// I:1800 (MONETcommon#17): a slew still running after 600 s is software error 16#40 and the slew is dropped. The time seam divides every
// timeout by 1000, so the 600 s are 0.6 s; the mock move takes far longer.
METHOD PRIVATE Slew_Times_Out_After_600_Seconds
VAR_INST
	rig			: FB_IagRig;
	nStep		: INT;
	nCycles		: UINT;
	sTest		: STRING(80);
END_VAR
TEST('Slew_Times_Out_After_600_Seconds');
sTest := 'Slew_Times_Out_After_600_Seconds: ';
IF nStep >= 90 THEN
	RETURN;
END_IF
rig.Scan();
nCycles := nCycles + 1;
CASE nStep OF
0:	// wait for the clock, then power on
	IF rig.ClockValid THEN
		rig.fbTel.Init();
		nStep := 10;
		nCycles := 0;
	ELSIF nCycles > 2000 THEN
		AssertTrue(Condition := FALSE, Message := 'the astronomical clock never became valid');
		F_Note(bFailed := TRUE, sText := CONCAT(sTest, 'the astronomical clock never became valid'));
		rig.SetTimeDivisor(nValue := 1);
		nStep := 99;
		TEST_FINISHED();
	END_IF
10:	IF rig.Online THEN
		rig.SetMoveScans(nScans := 60000);
		rig.SetTimeDivisor(nValue := 1000);
		rig.fbTel.Slew(fAzimuth := 180.0, fAltitude := 45.0);
		nStep := 20;
		nCycles := 0;
	ELSIF nCycles > 1500 THEN
		AssertTrue(Condition := FALSE, Message := 'the mock telescope did not reach READY_STATE 1.0');
		F_Note(bFailed := TRUE, sText := CONCAT(sTest, 'the mock telescope did not reach READY_STATE 1.0'));
		rig.SetTimeDivisor(nValue := 1);
		nStep := 99;
		TEST_FINISHED();
	END_IF
20:
	IF rig.fbTel.bError THEN
		AssertTrue(Condition := rig.fbTel.bSoftwareError AND rig.fbTel.nSoftwareErrorID = 16#40, Message := 'the slew timeout is software error 16#40');
		F_Note(bFailed := NOT (rig.fbTel.bSoftwareError AND rig.fbTel.nSoftwareErrorID = 16#40), sText := CONCAT(sTest, 'the slew timeout is software error 16#40'));
		AssertTrue(Condition := NOT rig.fbTel.bSlewActive, Message := 'the slew is dropped');
		F_Note(bFailed := NOT (NOT rig.fbTel.bSlewActive), sText := CONCAT(sTest, 'the slew is dropped'));
		rig.SetTimeDivisor(nValue := 1);
		nStep := 99;
		TEST_FINISHED();
	ELSIF nCycles > 3000 THEN
		AssertTrue(Condition := FALSE, Message := 'the slew never timed out');
		F_Note(bFailed := TRUE, sText := CONCAT(sTest, 'the slew never timed out'));
		rig.SetTimeDivisor(nValue := 1);
		nStep := 99;
		TEST_FINISHED();
	END_IF
END_CASE
END_METHOD

// I:466, 491-496: an online telescope without a command for 12 h parks itself (tonPowerTimeout). The time seam divides by 1000000, so the
// 12 h are 43 ms.
METHOD PRIVATE Idle_Telescope_Parks_After_12_Hours
VAR_INST
	rig			: FB_IagRig;
	nStep		: INT;
	nCycles		: UINT;
	sTest		: STRING(80);
END_VAR
TEST('Idle_Telescope_Parks_After_12_Hours');
sTest := 'Idle_Telescope_Parks_After_12_Hours: ';
IF nStep >= 90 THEN
	RETURN;
END_IF
rig.Scan();
nCycles := nCycles + 1;
CASE nStep OF
0:	// wait for the clock, then power on
	IF rig.ClockValid THEN
		rig.fbTel.Init();
		nStep := 10;
		nCycles := 0;
	ELSIF nCycles > 2000 THEN
		AssertTrue(Condition := FALSE, Message := 'the astronomical clock never became valid');
		F_Note(bFailed := TRUE, sText := CONCAT(sTest, 'the astronomical clock never became valid'));
		rig.SetTimeDivisor(nValue := 1);
		nStep := 99;
		TEST_FINISHED();
	END_IF
10:	IF rig.Online THEN
		rig.SetTimeDivisor(nValue := 1000000);
		nStep := 20;
		nCycles := 0;
	ELSIF nCycles > 1500 THEN
		AssertTrue(Condition := FALSE, Message := 'the mock telescope did not reach READY_STATE 1.0');
		F_Note(bFailed := TRUE, sText := CONCAT(sTest, 'the mock telescope did not reach READY_STATE 1.0'));
		rig.SetTimeDivisor(nValue := 1);
		nStep := 99;
		TEST_FINISHED();
	END_IF
20:
	IF rig.fbTel.bParkActive OR rig.fbTel.bIsParked THEN
		rig.SetTimeDivisor(nValue := 1);
		AssertTrue(Condition := rig.fbTel.bParkActive OR rig.fbTel.bIsParked, Message := 'the idle telescope parked itself');
		F_Note(bFailed := NOT (rig.fbTel.bParkActive OR rig.fbTel.bIsParked), sText := CONCAT(sTest, 'the idle telescope parked itself'));
		nStep := 99;
		TEST_FINISHED();
	ELSIF nCycles > 3000 THEN
		AssertTrue(Condition := FALSE, Message := 'the idle telescope never parked');
		F_Note(bFailed := TRUE, sText := CONCAT(sTest, 'the idle telescope never parked'));
		rig.SetTimeDivisor(nValue := 1);
		nStep := 99;
		TEST_FINISHED();
	END_IF
END_CASE
END_METHOD

END_FUNCTION_BLOCK

// ---- POUs/IagParkDuringPowerOn_Tests.TcPOU
// Characterization of FB_TelescopeControl (IAG50cm) for a park or a stop that arrives during the power-on, on mock axes (plan step 2,
// IAG50cmTests README). These tests pin what the code does today, with the line of the behaviour in a comment; they are not a
// specification. Every test owns a rig and runs over many PLC cycles (VAR_INST of the method, one Scan() per cycle). Failed checks
// are also noted in GVL_Diag.sFailures (printed by Run-Tests.ps1).
FUNCTION_BLOCK IagParkDuringPowerOn_Tests EXTENDS TcUnit.FB_TestSuite
VAR
END_VAR

Park_During_PowerOn_Aborts_The_Startup_And_Parks();
Stop_During_PowerOn_Aborts_The_Startup();
AxesOff_Park_After_Stopped_Startup_Reports_Parked();
AxesOff_Park_With_Slow_Covers_Reports_Parking_Then_Parked();
Stop_During_AxesOff_Park_Does_Not_Cancel_It();
AxesOff_Park_Gives_Up_When_The_Covers_Do_Not_Close();
Park_In_The_Sweep_Parks_In_Place();
Park_After_Stage_100_Still_Moves_To_The_Park_Position();

// I:529-541 (IAG50cm#109): a park that arrives while the power-on runs outranks it, like a stop: the startup is aborted, the
// covers the power-on opened are closed again and the telescope ends parked, never ready (READY_STATE does not reach 1.0).
// In the covers phase the axes are still off, so the park takes the axes-off path (#54, #110): covers closed, dome parked,
// the mount is not moved, READY_STATE 0.0 and bIsParked is TRUE with bParkedInPlace (#187). Decision 3 of the plan: as MONET (MONETcommon#87).
METHOD PRIVATE Park_During_PowerOn_Aborts_The_Startup_And_Parks
VAR_INST
	rig			: FB_IagRig;
	nStep		: INT;
	nCycles		: UINT;
	sTest		: STRING(80);
END_VAR
TEST('Park_During_PowerOn_Aborts_The_Startup_And_Parks');
sTest := 'Park_During_PowerOn_Aborts_The_Startup_And_Parks: ';
IF nStep >= 90 THEN
	RETURN;
END_IF
rig.Scan();
nCycles := nCycles + 1;
CASE nStep OF
0:	// wait for the clock, then power on
	IF rig.ClockValid THEN
		rig.fbTel.Init();
		nStep := 10;
		nCycles := 0;
	ELSIF nCycles > 2000 THEN
		AssertTrue(Condition := FALSE, Message := 'the astronomical clock never became valid');
		F_Note(bFailed := TRUE, sText := CONCAT(sTest, 'the astronomical clock never became valid'));
		nStep := 99;
		TEST_FINISHED();
	END_IF
10:	// the power-on has commanded the covers: park now
	IF rig.fbCovers.nOpenCalls >= 1 THEN
		rig.fbTel.Park();
		nStep := 20;
		nCycles := 0;
	ELSIF nCycles > 300 THEN
		AssertTrue(Condition := FALSE, Message := 'the power-on never commanded the covers');
		F_Note(bFailed := TRUE, sText := CONCAT(sTest, 'the power-on never commanded the covers'));
		nStep := 99;
		TEST_FINISHED();
	END_IF
20:	// the power-on is aborted at once, the covers are commanded closed
	IF nCycles = 3 THEN
		AssertTrue(Condition := NOT rig.fbTel.bPowerActive, Message := 'the power-on is aborted');
		F_Note(bFailed := (rig.fbTel.bPowerActive), sText := CONCAT(sTest, 'the power-on is aborted'));
		nStep := 30;
		nCycles := 0;
	END_IF
30:	// the park finishes (READY_STATE 0.0, the axes were off: bIsParked TRUE with bParkedInPlace, #187), the startup never does
	AssertFalse(Condition := rig.Online, Message := 'the startup went on to the end');
	F_Note(bFailed := (rig.Online), sText := CONCAT(sTest, 'the startup went on to the end'));
	IF rig.fbTel.ReadyState = 0.0 THEN
		AssertTrue(Condition := rig.fbCovers.nCloseCalls >= 1, Message := 'the covers were closed');
		F_Note(bFailed := NOT (rig.fbCovers.nCloseCalls >= 1), sText := CONCAT(sTest, 'the covers were closed'));
		AssertTrue(Condition := rig.fbTel.bIsParked, Message := 'bIsParked is TRUE (#187)');
		F_Note(bFailed := NOT (rig.fbTel.bIsParked), sText := CONCAT(sTest, 'bIsParked is TRUE (#187)'));
		AssertTrue(Condition := rig.fbTel.bParkedInPlace, Message := 'bParkedInPlace is TRUE, the mount was not moved');
		F_Note(bFailed := NOT (rig.fbTel.bParkedInPlace), sText := CONCAT(sTest, 'bParkedInPlace is TRUE, the mount was not moved'));
		nStep := 99;
		TEST_FINISHED();
	ELSIF nCycles > 1500 THEN
		AssertTrue(Condition := FALSE, Message := 'the telescope did not park');
		F_Note(bFailed := TRUE, sText := CONCAT(sTest, 'the telescope did not park'));
		nStep := 99;
		TEST_FINISHED();
	END_IF
END_CASE
END_METHOD

// I:501-526 (#27): an explicit stop outranks the power-on: the startup is aborted (READY_STATE -2.0), nothing is parked and the
// covers the power-on opened stay open.
METHOD PRIVATE Stop_During_PowerOn_Aborts_The_Startup
VAR_INST
	rig			: FB_IagRig;
	nStep		: INT;
	nCycles		: UINT;
	sTest		: STRING(80);
END_VAR
TEST('Stop_During_PowerOn_Aborts_The_Startup');
sTest := 'Stop_During_PowerOn_Aborts_The_Startup: ';
IF nStep >= 90 THEN
	RETURN;
END_IF
rig.Scan();
nCycles := nCycles + 1;
CASE nStep OF
0:	// wait for the clock, then power on
	IF rig.ClockValid THEN
		rig.fbTel.Init();
		nStep := 10;
		nCycles := 0;
	ELSIF nCycles > 2000 THEN
		AssertTrue(Condition := FALSE, Message := 'the astronomical clock never became valid');
		F_Note(bFailed := TRUE, sText := CONCAT(sTest, 'the astronomical clock never became valid'));
		nStep := 99;
		TEST_FINISHED();
	END_IF
10:	// the power-on has commanded the covers: stop now
	IF rig.fbCovers.nOpenCalls >= 1 THEN
		rig.fbTel.Stop();
		nStep := 20;
		nCycles := 0;
	ELSIF nCycles > 300 THEN
		AssertTrue(Condition := FALSE, Message := 'the power-on never commanded the covers');
		F_Note(bFailed := TRUE, sText := CONCAT(sTest, 'the power-on never commanded the covers'));
		nStep := 99;
		TEST_FINISHED();
	END_IF
20:	// wait until the stop has settled
	IF NOT rig.fbTel.bStopActive AND rig.fbTel.bStopped AND nCycles > 5 THEN
		AssertFalse(Condition := rig.fbTel.bPowerActive, Message := 'the power-on request is dropped');
		F_Note(bFailed := (rig.fbTel.bPowerActive), sText := CONCAT(sTest, 'the power-on request is dropped'));
		AssertFalse(Condition := rig.fbTel.bParkActive OR rig.fbTel.bIsParked, Message := 'the stop does not park');
		F_Note(bFailed := (rig.fbTel.bParkActive OR rig.fbTel.bIsParked), sText := CONCAT(sTest, 'the stop does not park'));
		AssertTrue(Condition := rig.fbTel.ReadyState = -2.0, Message := 'READY_STATE is -2.0 (startup aborted)');
		F_Note(bFailed := NOT (rig.fbTel.ReadyState = -2.0), sText := CONCAT(sTest, 'READY_STATE is -2.0 (startup aborted)'));
		AssertTrue(Condition := rig.fbCovers.nCloseCalls = 0 AND rig.fbCovers.bOpened, Message := 'the covers stay open');
		F_Note(bFailed := NOT (rig.fbCovers.nCloseCalls = 0 AND rig.fbCovers.bOpened), sText := CONCAT(sTest, 'the covers stay open'));
		nStep := 99;
		TEST_FINISHED();
	ELSIF nCycles > 400 THEN
		AssertTrue(Condition := FALSE, Message := 'the stop did not settle');
		F_Note(bFailed := TRUE, sText := CONCAT(sTest, 'the stop did not settle'));
		nStep := 99;
		TEST_FINISHED();
	END_IF
END_CASE
END_METHOD

// IAG50cm#110: after a stopped startup (-2) a park with the axes off closes the covers and parks the dome, the mount is not moved.
// READY_STATE leaves -2 for 0.0 and bIsParked becomes TRUE with bParkedInPlace (#187); a new power-on clears both.
METHOD PRIVATE AxesOff_Park_After_Stopped_Startup_Reports_Parked
VAR_INST
	rig			: FB_IagRig;
	nStep		: INT;
	nCycles		: UINT;
	sTest		: STRING(80);
END_VAR
TEST('AxesOff_Park_After_Stopped_Startup_Reports_Parked');
sTest := 'AxesOff_Park_After_Stopped_Startup_Reports_Parked: ';
IF nStep >= 90 THEN
	RETURN;
END_IF
rig.Scan();
nCycles := nCycles + 1;
CASE nStep OF
0:	// wait for the clock, then power on
	IF rig.ClockValid THEN
		rig.fbTel.Init();
		nStep := 10;
		nCycles := 0;
	ELSIF nCycles > 2000 THEN
		AssertTrue(Condition := FALSE, Message := 'the astronomical clock never became valid');
		F_Note(bFailed := TRUE, sText := CONCAT(sTest, 'the astronomical clock never became valid'));
		nStep := 99;
		TEST_FINISHED();
	END_IF
10:	// the power-on has commanded the covers: stop now
	IF rig.fbCovers.nOpenCalls >= 1 THEN
		rig.fbTel.Stop();
		nStep := 20;
		nCycles := 0;
	ELSIF nCycles > 300 THEN
		AssertTrue(Condition := FALSE, Message := 'the power-on never commanded the covers');
		F_Note(bFailed := TRUE, sText := CONCAT(sTest, 'the power-on never commanded the covers'));
		nStep := 99;
		TEST_FINISHED();
	END_IF
20:	// the stop has settled: -2, then park with the axes off
	IF NOT rig.fbTel.bStopActive AND rig.fbTel.bStopped AND nCycles > 5 THEN
		AssertTrue(Condition := rig.fbTel.ReadyState = -2.0, Message := 'READY_STATE is -2.0 after the stop');
		F_Note(bFailed := NOT (rig.fbTel.ReadyState = -2.0), sText := CONCAT(sTest, 'READY_STATE is -2.0 after the stop'));
		rig.fbTel.Park();
		nStep := 30;
		nCycles := 0;
	ELSIF nCycles > 400 THEN
		AssertTrue(Condition := FALSE, Message := 'the stop did not settle');
		F_Note(bFailed := TRUE, sText := CONCAT(sTest, 'the stop did not settle'));
		nStep := 99;
		TEST_FINISHED();
	END_IF
30:	// the covers close, READY_STATE becomes 0.0, bIsParked is TRUE (#187)
	IF rig.fbTel.ReadyState = 0.0 THEN
		AssertTrue(Condition := rig.fbCovers.nCloseCalls >= 1, Message := 'the covers were closed');
		F_Note(bFailed := NOT (rig.fbCovers.nCloseCalls >= 1), sText := CONCAT(sTest, 'the covers were closed'));
		AssertTrue(Condition := rig.fbTel.bIsParked, Message := 'bIsParked is TRUE (#187)');
		F_Note(bFailed := NOT (rig.fbTel.bIsParked), sText := CONCAT(sTest, 'bIsParked is TRUE (#187)'));
		AssertTrue(Condition := rig.fbTel.bParkedInPlace, Message := 'bParkedInPlace is TRUE, the mount was not moved');
		F_Note(bFailed := NOT (rig.fbTel.bParkedInPlace), sText := CONCAT(sTest, 'bParkedInPlace is TRUE, the mount was not moved'));
		rig.fbTel.Init();
		nStep := 40;
		nCycles := 0;
	ELSIF nCycles > 400 THEN
		AssertTrue(Condition := FALSE, Message := 'READY_STATE did not reach 0.0');
		F_Note(bFailed := TRUE, sText := CONCAT(sTest, 'READY_STATE did not reach 0.0'));
		nStep := 99;
		TEST_FINISHED();
	END_IF
40:	// a new power-on ends the covered state
	IF rig.fbTel.ReadyState > 0.0 THEN
		nStep := 99;
		TEST_FINISHED();
	ELSIF nCycles > 400 THEN
		AssertTrue(Condition := FALSE, Message := 'the new power-on did not leave READY_STATE 0.0');
		F_Note(bFailed := TRUE, sText := CONCAT(sTest, 'the new power-on did not leave READY_STATE 0.0'));
		nStep := 99;
		TEST_FINISHED();
	END_IF
END_CASE
END_METHOD

// IAG50cm#187: an axes-off park whose covers close slowly reports READY_STATE 0.3 and bIsParked FALSE while they are open, and
// parked in place (READY_STATE 0.0, bIsParked and bParkedInPlace TRUE) once they are closed. The covers mock holds the close.
METHOD PRIVATE AxesOff_Park_With_Slow_Covers_Reports_Parking_Then_Parked
VAR_INST
	rig			: FB_IagRig;
	nStep		: INT;
	nCycles		: UINT;
	sTest		: STRING(80);
END_VAR
TEST('AxesOff_Park_With_Slow_Covers_Reports_Parking_Then_Parked');
sTest := 'AxesOff_Park_With_Slow_Covers_Reports_Parking_Then_Parked: ';
IF nStep >= 90 THEN
	RETURN;
END_IF
rig.Scan();
nCycles := nCycles + 1;
CASE nStep OF
0:	// wait for the clock, then power on
	IF rig.ClockValid THEN
		rig.fbTel.Init();
		nStep := 10;
		nCycles := 0;
	ELSIF nCycles > 2000 THEN
		AssertTrue(Condition := FALSE, Message := 'the astronomical clock never became valid');
		F_Note(bFailed := TRUE, sText := CONCAT(sTest, 'the astronomical clock never became valid'));
		nStep := 99;
		TEST_FINISHED();
	END_IF
10:	// the power-on has commanded the covers: stop now
	IF rig.fbCovers.nOpenCalls >= 1 THEN
		rig.fbTel.Stop();
		nStep := 20;
		nCycles := 0;
	ELSIF nCycles > 300 THEN
		AssertTrue(Condition := FALSE, Message := 'the power-on never commanded the covers');
		F_Note(bFailed := TRUE, sText := CONCAT(sTest, 'the power-on never commanded the covers'));
		nStep := 99;
		TEST_FINISHED();
	END_IF
20:	// the stop has settled: the covers now close slowly, park with the axes off
	IF NOT rig.fbTel.bStopActive AND rig.fbTel.bStopped AND nCycles > 5 THEN
		rig.fbCovers.HoldClose(bHold := TRUE);
		rig.fbTel.Park();
		nStep := 30;
		nCycles := 0;
	ELSIF nCycles > 400 THEN
		AssertTrue(Condition := FALSE, Message := 'the stop did not settle');
		F_Note(bFailed := TRUE, sText := CONCAT(sTest, 'the stop did not settle'));
		nStep := 99;
		TEST_FINISHED();
	END_IF
30:	// the covers were commanded but are not closed: 0.3 (parking), not parked, not 0 and not -2
	IF rig.fbCovers.nCloseCalls >= 1 AND nCycles > 20 THEN
		AssertTrue(Condition := rig.fbTel.ReadyState = 0.3, Message := 'READY_STATE is 0.3 while the covers close (#187)');
		F_Note(bFailed := NOT (rig.fbTel.ReadyState = 0.3), sText := CONCAT(sTest, 'READY_STATE is 0.3 while the covers close (#187)'));
		AssertTrue(Condition := NOT rig.fbTel.bIsParked, Message := 'bIsParked stays FALSE until the covers are closed');
		F_Note(bFailed := NOT (NOT rig.fbTel.bIsParked), sText := CONCAT(sTest, 'bIsParked stays FALSE until the covers are closed'));
		AssertTrue(Condition := rig.fbTel.bSafeParked, Message := 'the axes-off park is pending');
		F_Note(bFailed := NOT (rig.fbTel.bSafeParked), sText := CONCAT(sTest, 'the axes-off park is pending'));
		rig.fbCovers.FinishClose();
		nStep := 40;
		nCycles := 0;
	ELSIF nCycles > 400 THEN
		AssertTrue(Condition := FALSE, Message := 'the covers were never commanded to close');
		F_Note(bFailed := TRUE, sText := CONCAT(sTest, 'the covers were never commanded to close'));
		nStep := 99;
		TEST_FINISHED();
	END_IF
40:	// the covers closed: parked in place
	IF rig.fbTel.ReadyState = 0.0 THEN
		AssertTrue(Condition := rig.fbTel.bIsParked, Message := 'bIsParked is TRUE once the covers are closed (#187)');
		F_Note(bFailed := NOT (rig.fbTel.bIsParked), sText := CONCAT(sTest, 'bIsParked is TRUE once the covers are closed (#187)'));
		AssertTrue(Condition := rig.fbTel.bParkedInPlace, Message := 'bParkedInPlace is TRUE, the mount was not moved');
		F_Note(bFailed := NOT (rig.fbTel.bParkedInPlace), sText := CONCAT(sTest, 'bParkedInPlace is TRUE, the mount was not moved'));
		AssertTrue(Condition := NOT rig.fbTel.bSafeParked, Message := 'the axes-off park is finished');
		F_Note(bFailed := NOT (NOT rig.fbTel.bSafeParked), sText := CONCAT(sTest, 'the axes-off park is finished'));
		nStep := 99;
		TEST_FINISHED();
	ELSIF nCycles > 400 THEN
		AssertTrue(Condition := FALSE, Message := 'READY_STATE did not reach 0.0 after the covers closed');
		F_Note(bFailed := TRUE, sText := CONCAT(sTest, 'READY_STATE did not reach 0.0 after the covers closed'));
		nStep := 99;
		TEST_FINISHED();
	END_IF
END_CASE
END_METHOD

// IAG50cm#196: a stop during the axes-off park (covers closing) is ignored and logged ('Stop ignored'): the park goes on and ends parked in place.
METHOD PRIVATE Stop_During_AxesOff_Park_Does_Not_Cancel_It
VAR_INST
	rig			: FB_IagRig;
	nStep		: INT;
	nCycles		: UINT;
	sTest		: STRING(80);
END_VAR
TEST('Stop_During_AxesOff_Park_Does_Not_Cancel_It');
sTest := 'Stop_During_AxesOff_Park_Does_Not_Cancel_It: ';
IF nStep >= 90 THEN
	RETURN;
END_IF
rig.Scan();
nCycles := nCycles + 1;
CASE nStep OF
0:	// wait for the clock, then power on
	IF rig.ClockValid THEN
		rig.fbTel.Init();
		nStep := 10;
		nCycles := 0;
	ELSIF nCycles > 2000 THEN
		AssertTrue(Condition := FALSE, Message := 'the astronomical clock never became valid');
		F_Note(bFailed := TRUE, sText := CONCAT(sTest, 'the astronomical clock never became valid'));
		nStep := 99;
		TEST_FINISHED();
	END_IF
10:	// the power-on has commanded the covers: stop now
	IF rig.fbCovers.nOpenCalls >= 1 THEN
		rig.fbTel.Stop();
		nStep := 20;
		nCycles := 0;
	ELSIF nCycles > 300 THEN
		AssertTrue(Condition := FALSE, Message := 'the power-on never commanded the covers');
		F_Note(bFailed := TRUE, sText := CONCAT(sTest, 'the power-on never commanded the covers'));
		nStep := 99;
		TEST_FINISHED();
	END_IF
20:	// the stop has settled: the covers now close slowly, park with the axes off
	IF NOT rig.fbTel.bStopActive AND rig.fbTel.bStopped AND nCycles > 5 THEN
		rig.fbCovers.HoldClose(bHold := TRUE);
		rig.fbTel.Park();
		nStep := 30;
		nCycles := 0;
	ELSIF nCycles > 400 THEN
		AssertTrue(Condition := FALSE, Message := 'the stop did not settle');
		F_Note(bFailed := TRUE, sText := CONCAT(sTest, 'the stop did not settle'));
		nStep := 99;
		TEST_FINISHED();
	END_IF
30:	// the covers were commanded but are not closed: 0.3 (parking), not parked, not 0 and not -2
	IF rig.fbCovers.nCloseCalls >= 1 AND nCycles > 20 THEN
		AssertTrue(Condition := rig.fbTel.ReadyState = 0.3, Message := 'READY_STATE is 0.3 while the covers close (#187)');
		F_Note(bFailed := NOT (rig.fbTel.ReadyState = 0.3), sText := CONCAT(sTest, 'READY_STATE is 0.3 while the covers close (#187)'));
		AssertTrue(Condition := NOT rig.fbTel.bIsParked, Message := 'bIsParked stays FALSE until the covers are closed');
		F_Note(bFailed := NOT (NOT rig.fbTel.bIsParked), sText := CONCAT(sTest, 'bIsParked stays FALSE until the covers are closed'));
		AssertTrue(Condition := rig.fbTel.bSafeParked, Message := 'the axes-off park is pending');
		F_Note(bFailed := NOT (rig.fbTel.bSafeParked), sText := CONCAT(sTest, 'the axes-off park is pending'));
		rig.fbTel.Stop();
		nStep := 35;
		nCycles := 0;
	ELSIF nCycles > 400 THEN
		AssertTrue(Condition := FALSE, Message := 'the covers were never commanded to close');
		F_Note(bFailed := TRUE, sText := CONCAT(sTest, 'the covers were never commanded to close'));
		nStep := 99;
		TEST_FINISHED();
	END_IF
35:	// the stop has settled: the park was not cancelled
	IF NOT rig.fbTel.bStopActive AND nCycles > 5 THEN
		AssertTrue(Condition := rig.fbTel.bSafeParked, Message := 'the stop does not cancel the axes-off park (#196)');
		F_Note(bFailed := NOT (rig.fbTel.bSafeParked), sText := CONCAT(sTest, 'the stop does not cancel the axes-off park (#196)'));
		AssertTrue(Condition := rig.fbTel.ReadyState = 0.3, Message := 'READY_STATE stays 0.3 after the stop (#196)');
		F_Note(bFailed := NOT (rig.fbTel.ReadyState = 0.3), sText := CONCAT(sTest, 'READY_STATE stays 0.3 after the stop (#196)'));
		rig.fbCovers.FinishClose();
		nStep := 40;
		nCycles := 0;
	ELSIF nCycles > 400 THEN
		AssertTrue(Condition := FALSE, Message := 'the stop did not settle');
		F_Note(bFailed := TRUE, sText := CONCAT(sTest, 'the stop did not settle'));
		nStep := 99;
		TEST_FINISHED();
	END_IF
40:	// the covers closed: parked in place
	IF rig.fbTel.ReadyState = 0.0 THEN
		AssertTrue(Condition := rig.fbTel.bIsParked, Message := 'bIsParked is TRUE once the covers are closed (#187)');
		F_Note(bFailed := NOT (rig.fbTel.bIsParked), sText := CONCAT(sTest, 'bIsParked is TRUE once the covers are closed (#187)'));
		AssertTrue(Condition := rig.fbTel.bParkedInPlace, Message := 'bParkedInPlace is TRUE, the mount was not moved');
		F_Note(bFailed := NOT (rig.fbTel.bParkedInPlace), sText := CONCAT(sTest, 'bParkedInPlace is TRUE, the mount was not moved'));
		AssertTrue(Condition := NOT rig.fbTel.bSafeParked, Message := 'the axes-off park is finished');
		F_Note(bFailed := NOT (NOT rig.fbTel.bSafeParked), sText := CONCAT(sTest, 'the axes-off park is finished'));
		nStep := 99;
		TEST_FINISHED();
	ELSIF nCycles > 400 THEN
		AssertTrue(Condition := FALSE, Message := 'READY_STATE did not reach 0.0 after the covers closed');
		F_Note(bFailed := TRUE, sText := CONCAT(sTest, 'READY_STATE did not reach 0.0 after the covers closed'));
		nStep := 99;
		TEST_FINISHED();
	END_IF
END_CASE
END_METHOD

// IAG50cm#187: an axes-off park whose covers never close gives up after 120 s (the time seam divides by 1000): bSafeParked is dropped,
// READY_STATE is not 0.3 for ever and the telescope is never reported parked.
METHOD PRIVATE AxesOff_Park_Gives_Up_When_The_Covers_Do_Not_Close
VAR_INST
	rig			: FB_IagRig;
	nStep		: INT;
	nCycles		: UINT;
	sTest		: STRING(80);
END_VAR
TEST('AxesOff_Park_Gives_Up_When_The_Covers_Do_Not_Close');
sTest := 'AxesOff_Park_Gives_Up_When_The_Covers_Do_Not_Close: ';
IF nStep >= 90 THEN
	RETURN;
END_IF
rig.Scan();
nCycles := nCycles + 1;
CASE nStep OF
0:	// wait for the clock, then power on
	IF rig.ClockValid THEN
		rig.fbTel.Init();
		nStep := 10;
		nCycles := 0;
	ELSIF nCycles > 2000 THEN
		AssertTrue(Condition := FALSE, Message := 'the astronomical clock never became valid');
		F_Note(bFailed := TRUE, sText := CONCAT(sTest, 'the astronomical clock never became valid'));
		nStep := 99;
		TEST_FINISHED();
	END_IF
10:	// the power-on has commanded the covers: stop now
	IF rig.fbCovers.nOpenCalls >= 1 THEN
		rig.fbTel.Stop();
		nStep := 20;
		nCycles := 0;
	ELSIF nCycles > 300 THEN
		AssertTrue(Condition := FALSE, Message := 'the power-on never commanded the covers');
		F_Note(bFailed := TRUE, sText := CONCAT(sTest, 'the power-on never commanded the covers'));
		nStep := 99;
		TEST_FINISHED();
	END_IF
20:	// the stop has settled: the covers never close, park with the axes off; 120 s are 0.12 s
	IF NOT rig.fbTel.bStopActive AND rig.fbTel.bStopped AND nCycles > 5 THEN
		rig.fbCovers.HoldClose(bHold := TRUE);
		rig.SetTimeDivisor(nValue := 1000);
		rig.fbTel.Park();
		nStep := 30;
		nCycles := 0;
	ELSIF nCycles > 400 THEN
		AssertTrue(Condition := FALSE, Message := 'the stop did not settle');
		F_Note(bFailed := TRUE, sText := CONCAT(sTest, 'the stop did not settle'));
		rig.SetTimeDivisor(nValue := 1);
		nStep := 99;
		TEST_FINISHED();
	END_IF
30:	// after the give-up the park is no longer pending: not 0.3 for ever, and never reported parked
	IF NOT rig.fbTel.bSafeParked AND nCycles > 5 THEN
		rig.SetTimeDivisor(nValue := 1);
		AssertTrue(Condition := NOT rig.fbTel.bIsParked, Message := 'bIsParked stays FALSE, the covers did not close (#187)');
		F_Note(bFailed := NOT (NOT rig.fbTel.bIsParked), sText := CONCAT(sTest, 'bIsParked stays FALSE, the covers did not close (#187)'));
		AssertTrue(Condition := NOT rig.fbTel.bParkedInPlace, Message := 'bParkedInPlace stays FALSE');
		F_Note(bFailed := NOT (NOT rig.fbTel.bParkedInPlace), sText := CONCAT(sTest, 'bParkedInPlace stays FALSE'));
		AssertTrue(Condition := rig.fbTel.ReadyState <> 0.3, Message := 'READY_STATE leaves 0.3 after the give-up');
		F_Note(bFailed := NOT (rig.fbTel.ReadyState <> 0.3), sText := CONCAT(sTest, 'READY_STATE leaves 0.3 after the give-up'));
		nStep := 99;
		TEST_FINISHED();
	ELSIF nCycles > 3000 THEN
		AssertTrue(Condition := FALSE, Message := 'the axes-off park never gave up');
		F_Note(bFailed := TRUE, sText := CONCAT(sTest, 'the axes-off park never gave up'));
		rig.SetTimeDivisor(nValue := 1);
		nStep := 99;
		TEST_FINISHED();
	END_IF
END_CASE
END_METHOD

// IAG50cm#197 (T38 step 2): a park in the calibration sweep (power-on stage 40 and later) aborts the startup, the axes are on, so the park
// can neither be dispatched (bReady needs the completed power-on) nor take the axes-off path. It used to hang at READY_STATE 0.3 for good.
// Now the axes are stopped and switched off once at rest, and the park ends parked in place (axes off, covers closed, dome parked).
// The mock axes do not hold the sweep after a stop (the real FB_HomeHold does), so the sweep runs to its end here: the park must still end.
METHOD PRIVATE Park_In_The_Sweep_Parks_In_Place
VAR_INST
	rig			: FB_IagRig;
	nStep		: INT;
	nCycles		: UINT;
	sTest		: STRING(80);
END_VAR
TEST('Park_In_The_Sweep_Parks_In_Place');
sTest := 'Park_In_The_Sweep_Parks_In_Place: ';
IF nStep >= 90 THEN
	RETURN;
END_IF
rig.Scan();
nCycles := nCycles + 1;
IF nStep >= 20 THEN
	// the startup never completes, and the telescope is never ready
	IF rig.fbTel.ReadyState = 1.0 OR rig.Online THEN
		AssertTrue(Condition := FALSE, Message := 'the startup went on to the end');
		F_Note(bFailed := TRUE, sText := CONCAT(sTest, 'the startup went on to the end'));
		nStep := 99;
		TEST_FINISHED();
	END_IF
END_IF
CASE nStep OF
0:	// wait for the clock, then power on with a long calibration sweep
	IF rig.ClockValid THEN
		rig.SetHomeScans(nHa := 400, nDec := 400);
		rig.fbTel.Init();
		nStep := 10;
		nCycles := 0;
	ELSIF nCycles > 2000 THEN
		AssertTrue(Condition := FALSE, Message := 'the astronomical clock never became valid');
		F_Note(bFailed := TRUE, sText := CONCAT(sTest, 'the astronomical clock never became valid'));
		nStep := 99;
		TEST_FINISHED();
	END_IF
10:	// both axes are enabled and sweeping (power-on stage 40): park now
	IF rig.fbHa.bEnable AND rig.fbDec.bEnable AND NOT rig.fbHa.bCalibrated AND NOT rig.fbDec.bCalibrated THEN
		nStep := 15;
		nCycles := 0;
	ELSIF nCycles > 3000 THEN
		AssertTrue(Condition := FALSE, Message := 'the power-on never reached the sweep');
		F_Note(bFailed := TRUE, sText := CONCAT(sTest, 'the power-on never reached the sweep'));
		nStep := 99;
		TEST_FINISHED();
	END_IF
15:	// the mock axes are ready after a few scans and then sweep (400 scans): park in the middle of it
	IF nCycles >= 20 THEN
		rig.fbTel.Park();
		nStep := 20;
		nCycles := 0;
	END_IF
20:	// the power-on is aborted at once
	IF nCycles = 3 THEN
		AssertTrue(Condition := NOT rig.fbTel.bPowerActive, Message := 'the power-on is aborted');
		F_Note(bFailed := (rig.fbTel.bPowerActive), sText := CONCAT(sTest, 'the power-on is aborted'));
		nStep := 30;
		nCycles := 0;
	END_IF
30:	// it ends parked in place: no hang at 0.3
	IF rig.fbTel.ReadyState = 0.0 AND rig.fbTel.bIsParked THEN
		AssertTrue(Condition := NOT rig.fbHa.bEnable AND NOT rig.fbDec.bEnable, Message := 'both axes are switched off');
		F_Note(bFailed := NOT (NOT rig.fbHa.bEnable AND NOT rig.fbDec.bEnable), sText := CONCAT(sTest, 'both axes are switched off'));
		AssertTrue(Condition := rig.fbHa.nStopEdges >= 1 AND rig.fbDec.nStopEdges >= 1, Message := 'both axes were sent a stop (#197 A1)');
		F_Note(bFailed := NOT (rig.fbHa.nStopEdges >= 1 AND rig.fbDec.nStopEdges >= 1), sText := CONCAT(sTest, 'both axes were sent a stop (#197 A1)'));
		AssertTrue(Condition := rig.fbTel.bParkedInPlace, Message := 'bParkedInPlace is TRUE');
		F_Note(bFailed := NOT (rig.fbTel.bParkedInPlace), sText := CONCAT(sTest, 'bParkedInPlace is TRUE'));
		AssertTrue(Condition := rig.fbCovers.nCloseCalls >= 1, Message := 'the covers were closed');
		F_Note(bFailed := NOT (rig.fbCovers.nCloseCalls >= 1), sText := CONCAT(sTest, 'the covers were closed'));
		AssertFalse(Condition := rig.fbTel.bError, Message := 'no error');
		F_Note(bFailed := (rig.fbTel.bError), sText := CONCAT(sTest, 'no error'));
		AssertFalse(Condition := rig.fbTel.bParkActive, Message := 'the park request ended');
		F_Note(bFailed := (rig.fbTel.bParkActive), sText := CONCAT(sTest, 'the park request ended'));
		nStep := 99;
		TEST_FINISHED();
	ELSIF nCycles > 3000 THEN
		AssertTrue(Condition := FALSE, Message := 'the park hangs (READY_STATE stays 0.3)');
		F_Note(bFailed := TRUE, sText := CONCAT(sTest, 'the park hangs (READY_STATE stays 0.3)'));
		nStep := 99;
		TEST_FINISHED();
	END_IF
END_CASE
END_METHOD

// IAG50cm#197 regression: a park of a completed power-on (bIsPowered TRUE, ready) takes the normal path (the mount is driven to the park
// position), not the in-place path: bParkedInPlace stays FALSE.
METHOD PRIVATE Park_After_Stage_100_Still_Moves_To_The_Park_Position
VAR_INST
	rig			: FB_IagRig;
	nStep		: INT;
	nCycles		: UINT;
	sTest		: STRING(80);
END_VAR
TEST('Park_After_Stage_100_Still_Moves_To_The_Park_Position');
sTest := 'Park_After_Stage_100_Still_Moves_To_The_Park_Position: ';
IF nStep >= 90 THEN
	RETURN;
END_IF
rig.Scan();
nCycles := nCycles + 1;
CASE nStep OF
0:	// wait for the clock, then power on
	IF rig.ClockValid THEN
		rig.fbTel.Init();
		nStep := 10;
		nCycles := 0;
	ELSIF nCycles > 2000 THEN
		AssertTrue(Condition := FALSE, Message := 'the astronomical clock never became valid');
		F_Note(bFailed := TRUE, sText := CONCAT(sTest, 'the astronomical clock never became valid'));
		nStep := 99;
		TEST_FINISHED();
	END_IF
10:	// the startup is complete: park
	IF rig.Online THEN
		rig.fbTel.Park();
		nStep := 20;
		nCycles := 0;
	ELSIF nCycles > 3000 THEN
		AssertTrue(Condition := FALSE, Message := 'the power-on never completed');
		F_Note(bFailed := TRUE, sText := CONCAT(sTest, 'the power-on never completed'));
		nStep := 99;
		TEST_FINISHED();
	END_IF
20:	// the park ends
	IF rig.fbTel.ReadyState = 0.0 AND rig.fbTel.bIsParked THEN
		AssertFalse(Condition := rig.fbTel.bParkedInPlace, Message := 'a park of a ready telescope is not an in-place park');
		F_Note(bFailed := (rig.fbTel.bParkedInPlace), sText := CONCAT(sTest, 'a park of a ready telescope is not an in-place park'));
		AssertFalse(Condition := rig.fbTel.bError, Message := 'no error');
		F_Note(bFailed := (rig.fbTel.bError), sText := CONCAT(sTest, 'no error'));
		nStep := 99;
		TEST_FINISHED();
	ELSIF nCycles > 4000 THEN
		AssertTrue(Condition := FALSE, Message := 'the park did not finish');
		F_Note(bFailed := TRUE, sText := CONCAT(sTest, 'the park did not finish'));
		nStep := 99;
		TEST_FINISHED();
	END_IF
END_CASE
END_METHOD

END_FUNCTION_BLOCK

// ---- POUs/IagStopDuringPark_Tests.TcPOU
// IAG50cm#92: a stop during the HA stage of a park, on mock axes (IAG50cmTests README). Unlike the characterization suites this is
// a regression test of a defect: it FAILS until #92 is fixed. Every test owns a rig and runs over many PLC cycles (VAR_INST of the
// method, one Scan() per cycle). Failed checks are also noted in GVL_Diag.sFailures (printed by Run-Tests.ps1).
FUNCTION_BLOCK IagStopDuringPark_Tests EXTENDS TcUnit.FB_TestSuite
VAR
	fDecAtStop	: LREAL;		// Dec actual position when the stop was sent
END_VAR

Stop_Right_After_The_HA_Stage_Of_A_Park_Still_Stops_Dec();

// #92 (T18.4): the park moves HA home first, then commands the Dec move (MoveAxis -> fbAxis.MoveTo()). The NC reports InMotion a few
// cycles later (mock: SetStartScans), so for those scans both axes still report StandStill (bStopped). A stop in that window runs for one
// scan only: bStop is cleared at once (bStopped), the first scan of _StopTelescope only drops MoveAxis (CancelMove does not
// stop a move that was already started) and the axis stop (StopAxis) is never sent. The Dec move to home runs to the end.
// Expected: Dec is sent a stop and stays where it was. (A stop before the Dec command works: TCS_command passes stop and Dec never starts.)
// CI trace of the defect (TCS_command, bStop, bStopped, bPark, Dec MoveAxis, Dec InMotion): park 2, 0,1,1,1,0 -> stop 5, 0,1,0,0,0 -> no_command 0, 0,1,0,0,0
// -> then Dec InMotion for the rest of its 60 scan move with bStopped FALSE and no stop sent.
METHOD PRIVATE Stop_Right_After_The_HA_Stage_Of_A_Park_Still_Stops_Dec
VAR_INST
	rig			: FB_IagRig;
	nStep		: INT;
	nCycles		: UINT;
	bHaMoved	: BOOL;
	bSawStop	: BOOL;
	sTest		: STRING(80);
END_VAR
TEST('Stop_Right_After_The_HA_Stage_Of_A_Park_Still_Stops_Dec');
sTest := 'Stop_Right_After_The_HA_Stage_Of_A_Park_Still_Stops_Dec: ';
IF nStep >= 90 THEN
	RETURN;
END_IF
rig.Scan();
nCycles := nCycles + 1;
CASE nStep OF
0:	// wait for the clock, then power on
	IF rig.ClockValid THEN
		rig.fbTel.Init();
		rig.SetStartScans(nScans := 3);
		nStep := 10;
		nCycles := 0;
	ELSIF nCycles > 2000 THEN
		AssertTrue(Condition := FALSE, Message := 'the astronomical clock never became valid');
		F_Note(bFailed := TRUE, sText := CONCAT(sTest, 'the astronomical clock never became valid'));
		nStep := 99;
		TEST_FINISHED();
	END_IF
10:	// ready: slew away from home to a point with an hour angle, so that the park moves HA first
	IF rig.Online THEN
		rig.fbTel.Slew(fAzimuth := 120.0, fAltitude := 40.0);
		nStep := 20;
		nCycles := 0;
	ELSIF nCycles > 1500 THEN
		AssertTrue(Condition := FALSE, Message := 'the mock telescope did not reach READY_STATE 1.0');
		F_Note(bFailed := TRUE, sText := CONCAT(sTest, 'the mock telescope did not reach READY_STATE 1.0'));
		nStep := 99;
		TEST_FINISHED();
	END_IF
20:	// the slew has finished and the mount stands still: park
	IF nCycles > 10 AND NOT rig.fbTel.bSlewActive AND rig.fbTel.bStopped AND rig.fbTel.TCS_command <> E_TCSCommand.slew THEN
		rig.fbTel.Park();
		nStep := 30;
		nCycles := 0;
	ELSIF nCycles > 600 THEN
		AssertTrue(Condition := FALSE, Message := 'the slew did not finish');
		F_Note(bFailed := TRUE, sText := CONCAT(sTest, 'the slew did not finish'));
		nStep := 99;
		TEST_FINISHED();
	END_IF
30:	// wait until HA has been moved by the park and the Dec move is commanded but the axis does not report InMotion yet: stop now
	IF rig.fbHa.MoveAxis THEN
		bHaMoved := TRUE;
	END_IF
	IF bHaMoved AND rig.fbDec.MoveAxis AND NOT rig.fbDec.fbAxis.InMotion AND rig.fbTel.bParkActive THEN
		fDecAtStop := rig.fbDec.fActualPosition;
		rig.fbTel.Stop();
		nStep := 40;
		nCycles := 0;
	ELSIF NOT rig.fbTel.bParkActive AND nCycles > 5 THEN
		AssertTrue(Condition := FALSE, Message := 'the park ended before the HA stage could be observed');
		F_Note(bFailed := TRUE, sText := CONCAT(sTest, 'the park ended before the HA stage could be observed'));
		nStep := 99;
		TEST_FINISHED();
	ELSIF nCycles > 600 THEN
		AssertTrue(Condition := FALSE, Message := 'the park never finished its HA stage');
		F_Note(bFailed := TRUE, sText := CONCAT(sTest, 'the park never finished its HA stage'));
		nStep := 99;
		TEST_FINISHED();
	END_IF
40:	// the mock Dec move takes 60 scans: look when it would have ended
	IF rig.fbTel.TCS_command = E_TCSCommand.stop THEN
		bSawStop := TRUE;
	END_IF
	IF nCycles >= 100 THEN
		AssertTrue(Condition := bSawStop, Message := 'the stop command ran (TCS_command passed stop)');
		F_Note(bFailed := NOT (bSawStop), sText := CONCAT(sTest, 'the stop command ran (TCS_command passed stop)'));
		AssertFalse(Condition := rig.fbTel.bParkActive, Message := 'the park is cancelled');
		F_Note(bFailed := (rig.fbTel.bParkActive), sText := CONCAT(sTest, 'the park is cancelled'));
		AssertTrue(Condition := rig.fbDec.nStopEdges >= 1, Message := 'Dec was sent an axis stop (the Dec move had started)');
		F_Note(bFailed := NOT (rig.fbDec.nStopEdges >= 1), sText := CONCAT(sTest, 'Dec was sent an axis stop (the Dec move had started)'));
		AssertTrue(Condition := rig.fbDec.fActualPosition = fDecAtStop, Message := 'Dec did not move to home after the stop');
		F_Note(bFailed := NOT (rig.fbDec.fActualPosition = fDecAtStop), sText := CONCAT(sTest, 'Dec did not move to home after the stop'));
		nStep := 99;
		TEST_FINISHED();
	END_IF
END_CASE
END_METHOD

END_FUNCTION_BLOCK

// ---- POUs/IagParkInLimit_Tests.TcPOU
// IAG50cm#84: a park requested while the mount stands inside the horizon limit homes out of the limit first and then parks
// (it used to starve against the safety block's automatic home). The mount is put in the limit by raising fHorizon above its
// elevation; the mock rig does not interpolate, so this tests the arbitration, not the real path altitude.
// Failed checks are also noted in GVL_Diag.sFailures (printed by Run-Tests.ps1).
FUNCTION_BLOCK IagParkInLimit_Tests EXTENDS TcUnit.FB_TestSuite
VAR
END_VAR

Park_Stopped_In_Limit_Homes_Then_Parks();
User_Stop_Cancels_The_Park_Waiting_For_The_Home();
Parked_With_Stale_Target_Below_Horizon_Raises_No_Horizon_Event();

// I:FB_TelescopeControl safety blocks, park branch (#84): home, then park; no stop, the covers close at the park.
METHOD PRIVATE Park_Stopped_In_Limit_Homes_Then_Parks
VAR_INST
	rig			: FB_IagRig;
	nStep		: INT;
	nCycles		: UINT;
	nStopsHa	: UINT;
	nStopsDec	: UINT;
	bHomeSeen	: BOOL;
	sTest		: STRING(80);
END_VAR
TEST('Park_Stopped_In_Limit_Homes_Then_Parks');
sTest := 'Park_Stopped_In_Limit_Homes_Then_Parks: ';
IF nStep >= 90 THEN
	RETURN;
END_IF
rig.Scan();
nCycles := nCycles + 1;
CASE nStep OF
0:	// wait for the clock, then power on
	IF rig.ClockValid THEN
		rig.fbTel.Init();
		nStep := 10;
		nCycles := 0;
	ELSIF nCycles > 2000 THEN
		AssertTrue(Condition := FALSE, Message := 'the astronomical clock never became valid');
		F_Note(bFailed := TRUE, sText := CONCAT(sTest, 'the astronomical clock never became valid'));
		nStep := 99;
		TEST_FINISHED();
	END_IF
10:	// wait until the startup has finished, then slew to 45 deg elevation
	IF rig.Online THEN
		rig.fbTel.Slew(fAzimuth := 180.0, fAltitude := 45.0);
		nStep := 15;
		nCycles := 0;
	ELSIF nCycles > 1500 THEN
		AssertTrue(Condition := FALSE, Message := 'the mock telescope did not reach READY_STATE 1.0');
		F_Note(bFailed := TRUE, sText := CONCAT(sTest, 'the mock telescope did not reach READY_STATE 1.0'));
		nStep := 99;
		TEST_FINISHED();
	END_IF
15:	// wait until the slew is done and the mount stands still
	IF NOT rig.fbTel.bSlewActive AND rig.fbTel.bStopped AND nCycles > 5 THEN
		nStopsHa := rig.fbHa.nStopEdges;
		nStopsDec := rig.fbDec.nStopEdges;
		// the mount now stands at 45 deg: raise the horizon limit above it and park (#84)
		rig.SetHorizon(fValue := 60.0);
		rig.fbTel.Park();
		nStep := 20;
		nCycles := 0;
	ELSIF nCycles > 800 THEN
		AssertTrue(Condition := FALSE, Message := 'the slew did not finish');
		F_Note(bFailed := TRUE, sText := CONCAT(sTest, 'the slew did not finish'));
		nStep := 99;
		TEST_FINISHED();
	END_IF
20:	// the home out of the limit runs first, the park follows
	bHomeSeen := bHomeSeen OR (rig.fbTel.bGoHomeActive AND rig.fbTel.bParkActive);
	IF rig.fbTel.bIsParked AND NOT rig.fbTel.bParkActive THEN
		AssertTrue(Condition := bHomeSeen, Message := 'the home ran while the park was pending');
		F_Note(bFailed := NOT (bHomeSeen), sText := CONCAT(sTest, 'the home ran while the park was pending'));
		AssertTrue(Condition := rig.fbHa.nStopEdges = nStopsHa AND rig.fbDec.nStopEdges = nStopsDec, Message := 'no stop was sent to the axes');
		F_Note(bFailed := NOT (rig.fbHa.nStopEdges = nStopsHa AND rig.fbDec.nStopEdges = nStopsDec), sText := CONCAT(sTest, 'no stop was sent to the axes'));
		AssertTrue(Condition := rig.fbCovers.nCloseCalls >= 1, Message := 'the covers were closed');
		F_Note(bFailed := NOT (rig.fbCovers.nCloseCalls >= 1), sText := CONCAT(sTest, 'the covers were closed'));
		nStep := 99;
		TEST_FINISHED();
	ELSIF nCycles > 2500 THEN
		AssertTrue(Condition := FALSE, Message := 'the park did not complete');
		F_Note(bFailed := TRUE, sText := CONCAT(sTest, 'the park did not complete'));
		nStep := 99;
		TEST_FINISHED();
	END_IF
END_CASE
END_METHOD

// #84: a user stop drops the pending park and its home; the park is not replayed.
METHOD PRIVATE User_Stop_Cancels_The_Park_Waiting_For_The_Home
VAR_INST
	rig			: FB_IagRig;
	nStep		: INT;
	nCycles		: UINT;
	nStopsHa	: UINT;
	nStopsDec	: UINT;
	bHomeSeen	: BOOL;
	sTest		: STRING(80);
END_VAR
TEST('User_Stop_Cancels_The_Park_Waiting_For_The_Home');
sTest := 'User_Stop_Cancels_The_Park_Waiting_For_The_Home: ';
IF nStep >= 90 THEN
	RETURN;
END_IF
rig.Scan();
nCycles := nCycles + 1;
CASE nStep OF
0:	// wait for the clock, then power on
	IF rig.ClockValid THEN
		rig.fbTel.Init();
		nStep := 10;
		nCycles := 0;
	ELSIF nCycles > 2000 THEN
		AssertTrue(Condition := FALSE, Message := 'the astronomical clock never became valid');
		F_Note(bFailed := TRUE, sText := CONCAT(sTest, 'the astronomical clock never became valid'));
		nStep := 99;
		TEST_FINISHED();
	END_IF
10:	// wait until the startup has finished, then slew to 45 deg elevation
	IF rig.Online THEN
		rig.fbTel.Slew(fAzimuth := 180.0, fAltitude := 45.0);
		nStep := 15;
		nCycles := 0;
	ELSIF nCycles > 1500 THEN
		AssertTrue(Condition := FALSE, Message := 'the mock telescope did not reach READY_STATE 1.0');
		F_Note(bFailed := TRUE, sText := CONCAT(sTest, 'the mock telescope did not reach READY_STATE 1.0'));
		nStep := 99;
		TEST_FINISHED();
	END_IF
15:	// wait until the slew is done and the mount stands still
	IF NOT rig.fbTel.bSlewActive AND rig.fbTel.bStopped AND nCycles > 5 THEN
		nStopsHa := rig.fbHa.nStopEdges;
		nStopsDec := rig.fbDec.nStopEdges;
		// the mount now stands at 45 deg: raise the horizon limit above it and park (#84)
		rig.SetHorizon(fValue := 60.0);
		rig.fbTel.Park();
		nStep := 20;
		nCycles := 0;
	ELSIF nCycles > 800 THEN
		AssertTrue(Condition := FALSE, Message := 'the slew did not finish');
		F_Note(bFailed := TRUE, sText := CONCAT(sTest, 'the slew did not finish'));
		nStep := 99;
		TEST_FINISHED();
	END_IF
20:	// the park waits for the home: stop
	IF rig.fbTel.bParkActive AND rig.fbTel.bGoHomeActive AND nCycles >= 3 THEN
		rig.fbTel.Stop();
		nStep := 30;
		nCycles := 0;
	ELSIF nCycles > 300 THEN
		AssertTrue(Condition := FALSE, Message := 'the park never waited for the home');
		F_Note(bFailed := TRUE, sText := CONCAT(sTest, 'the park never waited for the home'));
		nStep := 99;
		TEST_FINISHED();
	END_IF
30:	// the stop drops the park and the home; the park does not come back
	IF nCycles = 5 THEN
		AssertTrue(Condition := NOT rig.fbTel.bParkActive, Message := 'the stop cancelled the park');
		F_Note(bFailed := NOT (NOT rig.fbTel.bParkActive), sText := CONCAT(sTest, 'the stop cancelled the park'));
	END_IF
	IF nCycles > 400 THEN
		AssertTrue(Condition := NOT rig.fbTel.bParkActive AND NOT rig.fbTel.bIsParked, Message := 'the park did not replay after the stop');
		F_Note(bFailed := NOT (NOT rig.fbTel.bParkActive AND NOT rig.fbTel.bIsParked), sText := CONCAT(sTest, 'the park did not replay after the stop'));
		AssertTrue(Condition := rig.fbCovers.nCloseCalls = 0, Message := 'the covers stay open');
		F_Note(bFailed := NOT (rig.fbCovers.nCloseCalls = 0), sText := CONCAT(sTest, 'the covers stay open'));
		nStep := 99;
		TEST_FINISHED();
	END_IF
END_CASE
END_METHOD

// IAG50cm#127 (MONETcommon#94): the 'Target below safe horizon' event is only for a requested goto/slew. A parked telescope
// whose last target is below the horizon limit must not raise it.
METHOD PRIVATE Parked_With_Stale_Target_Below_Horizon_Raises_No_Horizon_Event
VAR_INST
	rig			: FB_IagRig;
	nStep		: INT;
	nCycles		: UINT;
	bEventSeen	: BOOL;
	sTest		: STRING(80);
END_VAR
TEST('Parked_With_Stale_Target_Below_Horizon_Raises_No_Horizon_Event');
sTest := 'Parked_With_Stale_Target_Below_Horizon_Raises_No_Horizon_Event: ';
IF nStep >= 90 THEN
	RETURN;
END_IF
rig.Scan();
nCycles := nCycles + 1;
CASE nStep OF
0:	// wait for the clock, then power on
	IF rig.ClockValid THEN
		rig.fbTel.Init();
		nStep := 10;
		nCycles := 0;
	ELSIF nCycles > 2000 THEN
		AssertTrue(Condition := FALSE, Message := 'the astronomical clock never became valid');
		F_Note(bFailed := TRUE, sText := CONCAT(sTest, 'the astronomical clock never became valid'));
		nStep := 99;
		TEST_FINISHED();
	END_IF
10:	// wait until the startup has finished, then slew to 45 deg elevation (the target the park leaves behind)
	IF rig.Online THEN
		rig.fbTel.Slew(fAzimuth := 180.0, fAltitude := 45.0);
		nStep := 15;
		nCycles := 0;
	ELSIF nCycles > 1500 THEN
		AssertTrue(Condition := FALSE, Message := 'the mock telescope did not reach READY_STATE 1.0');
		F_Note(bFailed := TRUE, sText := CONCAT(sTest, 'the mock telescope did not reach READY_STATE 1.0'));
		nStep := 99;
		TEST_FINISHED();
	END_IF
15:	// wait until the slew is done, then park
	IF NOT rig.fbTel.bSlew AND rig.fbTel.bStopped AND nCycles > 5 THEN
		rig.fbTel.Park();
		nStep := 20;
		nCycles := 0;
	ELSIF nCycles > 800 THEN
		AssertTrue(Condition := FALSE, Message := 'the slew did not finish');
		F_Note(bFailed := TRUE, sText := CONCAT(sTest, 'the slew did not finish'));
		nStep := 99;
		TEST_FINISHED();
	END_IF
20:	// wait until parked and no goto/slew is left, then put the stale target below the horizon limit
	IF rig.fbTel.bIsParked AND NOT rig.fbTel.bPark THEN
		AssertTrue(Condition := NOT rig.fbTel.bGoto AND NOT rig.fbTel.bSlew, Message := 'no goto/slew request is left after the park');
		F_Note(bFailed := NOT (NOT rig.fbTel.bGoto AND NOT rig.fbTel.bSlew), sText := CONCAT(sTest, 'no goto/slew request is left after the park'));
		rig.SetHorizon(fValue := 60.0);
		nStep := 30;
		nCycles := 0;
	ELSIF nCycles > 2500 THEN
		AssertTrue(Condition := FALSE, Message := 'the park did not complete');
		F_Note(bFailed := TRUE, sText := CONCAT(sTest, 'the park did not complete'));
		nStep := 99;
		TEST_FINISHED();
	END_IF
30:	// the event trigger is a one-scan pulse: sample every scan
	bEventSeen := bEventSeen OR rig.fbTel.rtrigHorizonError.Q;
	IF nCycles > 300 THEN
		AssertTrue(Condition := NOT bEventSeen, Message := 'no horizon event on a parked telescope');
		F_Note(bFailed := bEventSeen, sText := CONCAT(sTest, 'no horizon event on a parked telescope'));
		nStep := 99;
		TEST_FINISHED();
	END_IF
END_CASE
END_METHOD

END_FUNCTION_BLOCK

// ---- POUs/IagStuckStop_Tests.TcPOU
// IAG50cm#120: a stop transaction whose axis never reports Done, on mock axes (SetStopWithoutDone). Before the fix the
// transaction stayed open for good (bSettled FALSE) and held every home behind the stop. Same shape as IagStopDuringSlew_Tests:
// one rig per test, one Scan() per PLC cycle, a step that does not happen within its budget fails the test.
FUNCTION_BLOCK IagStuckStop_Tests EXTENDS TcUnit.FB_TestSuite
VAR
END_VAR

Stuck_Stop_At_Rest_Is_Released_After_The_Timeout();

// Slew, stop, and the moving axis never reports its stop Done. The axes are at rest at once, but the transaction stays
// open (bSettled FALSE) until the 30 s timeout (the time seam divides it by 100: 0.3 s); then it settles with no second stop,
// no error, and StopAxis of the axis is cleared so that the next stop gives a rising edge.
METHOD PRIVATE Stuck_Stop_At_Rest_Is_Released_After_The_Timeout
VAR_INST
	rig			: FB_IagRig;
	nStep		: INT;
	nCycles		: UINT;
	sTest		: STRING(80);
END_VAR
TEST('Stuck_Stop_At_Rest_Is_Released_After_The_Timeout');
sTest := 'Stuck_Stop_At_Rest_Is_Released_After_The_Timeout: ';
IF nStep >= 90 THEN
	RETURN;
END_IF
rig.Scan();
nCycles := nCycles + 1;
CASE nStep OF
0:	// wait for the clock, then power on
	IF rig.ClockValid THEN
		rig.fbTel.Init();
		nStep := 10;
		nCycles := 0;
	ELSIF nCycles > 2000 THEN
		AssertTrue(Condition := FALSE, Message := 'the astronomical clock never became valid');
		F_Note(bFailed := TRUE, sText := CONCAT(sTest, 'the astronomical clock never became valid'));
		nStep := 99;
		TEST_FINISHED();
	END_IF
10:	// wait until the startup has finished (READY_STATE 1.0), then slew with both mock stops losing their Done
	IF rig.Online THEN
		rig.SetStopWithoutDone(bHa := TRUE, bDec := TRUE);
		rig.SetTimeDivisor(nValue := 100);
		rig.fbTel.Slew(fAzimuth := 180.0, fAltitude := 45.0);
		nStep := 20;
		nCycles := 0;
	ELSIF nCycles > 1500 THEN
		AssertTrue(Condition := FALSE, Message := 'the mock telescope did not reach READY_STATE 1.0');
		F_Note(bFailed := TRUE, sText := CONCAT(sTest, 'the mock telescope did not reach READY_STATE 1.0'));
		nStep := 99;
		TEST_FINISHED();
	END_IF
20:	// wait until one axis is moving, let it run a few scans, then stop
	IF rig.fbHa.MoveAxis OR rig.fbDec.MoveAxis THEN
		IF nCycles >= 5 THEN
			rig.fbTel.Stop();
			nStep := 30;
			nCycles := 0;
		END_IF
	ELSIF nCycles > 300 THEN
		AssertTrue(Condition := FALSE, Message := 'the slew did not start an axis move');
		F_Note(bFailed := TRUE, sText := CONCAT(sTest, 'the slew did not start an axis move'));
		rig.SetTimeDivisor(nValue := 1);
		nStep := 99;
		TEST_FINISHED();
	END_IF
30:	// the stop has taken the axes to rest, but the transaction is still open: nothing has reported Done, so the stop is held (3A.2)
	IF rig.fbTel.bStopped AND nCycles > 3 THEN
		AssertFalse(Condition := rig.fbTel.bSettled, Message := 'not settled before the timeout: the axis never reported Done');
		F_Note(bFailed := rig.fbTel.bSettled, sText := CONCAT(sTest, 'not settled before the timeout: the axis never reported Done'));
		AssertTrue(Condition := rig.fbTel.bStopActive, Message := 'the stop is held until the transaction settles');
		F_Note(bFailed := NOT rig.fbTel.bStopActive, sText := CONCAT(sTest, 'the stop is held until the transaction settles'));
		nStep := 40;
		nCycles := 0;
	ELSIF nCycles > 400 THEN
		AssertTrue(Condition := FALSE, Message := 'the stop did not bring the axes to rest');
		F_Note(bFailed := TRUE, sText := CONCAT(sTest, 'the stop did not bring the axes to rest'));
		rig.SetTimeDivisor(nValue := 1);
		nStep := 99;
		TEST_FINISHED();
	END_IF
40:	// the timeout releases the transaction (0.3 s in the divided time)
	IF rig.fbTel.bSettled THEN
		AssertEquals_UINT(Expected := UINT#1, Actual := rig.fbHa.nStopEdges + rig.fbDec.nStopEdges, Message := 'one stop request in all, no second one after the timeout');
		F_Note(bFailed := (UINT#1) <> (rig.fbHa.nStopEdges + rig.fbDec.nStopEdges), sText := CONCAT(sTest, 'one stop request in all, no second one after the timeout'));
		AssertFalse(Condition := rig.fbTel.bError OR rig.fbTel.bSoftwareError, Message := 'no error: the release is not a fault');
		F_Note(bFailed := rig.fbTel.bError OR rig.fbTel.bSoftwareError, sText := CONCAT(sTest, 'no error: the release is not a fault'));
		AssertFalse(Condition := rig.fbHa.StopAxis OR rig.fbDec.StopAxis, Message := 'StopAxis cleared at the release');
		F_Note(bFailed := rig.fbHa.StopAxis OR rig.fbDec.StopAxis, sText := CONCAT(sTest, 'StopAxis cleared at the release'));
		rig.SetTimeDivisor(nValue := 1);
		nStep := 99;
		TEST_FINISHED();
	ELSIF nCycles > 3000 THEN
		AssertTrue(Condition := FALSE, Message := 'the stuck stop was never released');
		F_Note(bFailed := TRUE, sText := CONCAT(sTest, 'the stuck stop was never released'));
		rig.SetTimeDivisor(nValue := 1);
		nStep := 99;
		TEST_FINISHED();
	END_IF
END_CASE
END_METHOD

END_FUNCTION_BLOCK

// ---- POUs/IagCommandInputs_Tests.TcPOU
// The command inputs bStop/bPark/bPower/bReset of FB_TelescopeControl (IAG50cm) are edge-triggered like the methods and are never
// written by the block; the block works on the request latches bStopActive/bParkActive/bPowerActive/bResetActive.
// Plan: BROTLib specs/plans/2026-11-09-iag50cm-command-model-unification.md, steps 1a/1b. One rig per test, one Scan() per PLC cycle.
FUNCTION_BLOCK IagCommandInputs_Tests EXTENDS TcUnit.FB_TestSuite
VAR
END_VAR

Held_Stop_Input_Stops_Once();
Park_Input_Edge_Parks_Like_Park();
Stop_Method_And_Input_Edge_In_One_Scan_Count_Once();
Power_Input_Is_Not_Written_By_The_Block();
Held_Slew_Input_Starts_The_Slew_Once();
Slew_Input_Falling_Does_Not_Abort_The_Slew();
Slew_Method_And_Input_Edge_In_One_Scan_Count_Once();
Slew_Input_In_The_Scan_Of_A_New_Error_Is_Rejected();
Track_Method_And_Track_Input_In_One_Scan_Count_Once();

// A held stop input is one command: one stop transaction, never repeated, never cleared by the block (IAG50cm command model step 1a).
METHOD PRIVATE Held_Stop_Input_Stops_Once
VAR_INST
	rig			: FB_IagRig;
	nStep		: INT;
	nCycles		: UINT;
	nEdges		: UINT;
	sTest		: STRING(80);
END_VAR
TEST('Held_Stop_Input_Stops_Once');
sTest := 'Held_Stop_Input_Stops_Once: ';
IF nStep >= 90 THEN
	RETURN;
END_IF
rig.Scan();
nCycles := nCycles + 1;
CASE nStep OF
0:	// wait for the clock, then power on
	IF rig.ClockValid THEN
		rig.fbTel.Init();
		nStep := 10;
		nCycles := 0;
	ELSIF nCycles > 2000 THEN
		AssertTrue(Condition := FALSE, Message := 'the astronomical clock never became valid');
		F_Note(bFailed := TRUE, sText := CONCAT(sTest, 'the astronomical clock never became valid'));
		nStep := 99;
		TEST_FINISHED();
	END_IF
10:	// wait until the startup has finished (READY_STATE 1.0)
	IF rig.Online THEN
		rig.fbTel.Slew(fAzimuth := 180.0, fAltitude := 45.0);
		nStep := 20;
		nCycles := 0;
	ELSIF nCycles > 1500 THEN
		AssertTrue(Condition := FALSE, Message := 'the mock telescope did not reach READY_STATE 1.0');
		F_Note(bFailed := TRUE, sText := CONCAT(sTest, 'the mock telescope did not reach READY_STATE 1.0'));
		nStep := 99;
		TEST_FINISHED();
	END_IF
20:	// an axis is moving
	IF rig.fbHa.MoveAxis OR rig.fbDec.MoveAxis THEN
		nCycles := 0;
		nStep := 30;
	ELSIF nCycles > 300 THEN
		AssertTrue(Condition := FALSE, Message := 'the slew did not start an axis move');
		F_Note(bFailed := TRUE, sText := CONCAT(sTest, 'the slew did not start an axis move'));
		nStep := 99;
		TEST_FINISHED();
	END_IF
30:	// a few scans of motion, then hold the stop INPUT (an ADS write, not the method)
	IF nCycles >= 5 THEN
		rig.SetStopInput(TRUE);
		nStep := 40;
		nCycles := 0;
	END_IF
40:	// the stop has settled: note the stop edges, keep holding the input
	IF NOT rig.fbTel.bStopActive AND rig.fbTel.bStopped AND nCycles > 5 THEN
		nEdges := rig.fbHa.nStopEdges + rig.fbDec.nStopEdges;
		AssertTrue(Condition := nEdges = 1, Message := 'the held input sent one stop to the moving axis');
		F_Note(bFailed := NOT (nEdges = 1), sText := CONCAT(sTest, 'the held input sent one stop to the moving axis'));
		nStep := 50;
		nCycles := 0;
	ELSIF nCycles > 400 THEN
		AssertTrue(Condition := FALSE, Message := 'the stop did not settle');
		F_Note(bFailed := TRUE, sText := CONCAT(sTest, 'the stop did not settle'));
		nStep := 99;
		TEST_FINISHED();
	END_IF
50:	// 60 more scans with the input still TRUE: no second stop, the latch stays down, the input is not cleared
	IF nCycles >= 60 THEN
		AssertTrue(Condition := rig.fbHa.nStopEdges + rig.fbDec.nStopEdges = nEdges, Message := 'a held input is not a second stop');
		F_Note(bFailed := NOT (rig.fbHa.nStopEdges + rig.fbDec.nStopEdges = nEdges), sText := CONCAT(sTest, 'a held input is not a second stop'));
		AssertTrue(Condition := NOT rig.fbTel.bStopActive, Message := 'the stop latch stayed down');
		F_Note(bFailed := NOT (NOT rig.fbTel.bStopActive), sText := CONCAT(sTest, 'the stop latch stayed down'));
		AssertTrue(Condition := rig.fbTel.bStop, Message := 'the block did not clear the input');
		F_Note(bFailed := NOT (rig.fbTel.bStop), sText := CONCAT(sTest, 'the block did not clear the input'));
		AssertTrue(Condition := rig.fbFocus.nStop = 1, Message := 'one stop for the focus');
		F_Note(bFailed := NOT (rig.fbFocus.nStop = 1), sText := CONCAT(sTest, 'one stop for the focus'));
		nStep := 99;
		TEST_FINISHED();
	END_IF
END_CASE
END_METHOD

// A rising park input starts the park exactly like Park(); the finished park is not replayed from the held input.
METHOD PRIVATE Park_Input_Edge_Parks_Like_Park
VAR_INST
	rig			: FB_IagRig;
	nStep		: INT;
	nCycles		: UINT;
	nEdges		: UINT;
	sTest		: STRING(80);
END_VAR
TEST('Park_Input_Edge_Parks_Like_Park');
sTest := 'Park_Input_Edge_Parks_Like_Park: ';
IF nStep >= 90 THEN
	RETURN;
END_IF
rig.Scan();
nCycles := nCycles + 1;
CASE nStep OF
0:	// wait for the clock, then power on
	IF rig.ClockValid THEN
		rig.fbTel.Init();
		nStep := 10;
		nCycles := 0;
	ELSIF nCycles > 2000 THEN
		AssertTrue(Condition := FALSE, Message := 'the astronomical clock never became valid');
		F_Note(bFailed := TRUE, sText := CONCAT(sTest, 'the astronomical clock never became valid'));
		nStep := 99;
		TEST_FINISHED();
	END_IF
10:	// wait until the startup has finished (READY_STATE 1.0)
	IF rig.Online THEN
		rig.SetParkInput(TRUE);
		nStep := 20;
		nCycles := 0;
	ELSIF nCycles > 1500 THEN
		AssertTrue(Condition := FALSE, Message := 'the mock telescope did not reach READY_STATE 1.0');
		F_Note(bFailed := TRUE, sText := CONCAT(sTest, 'the mock telescope did not reach READY_STATE 1.0'));
		nStep := 99;
		TEST_FINISHED();
	END_IF
20:	// the edge starts the park, as Park() would
	IF rig.fbTel.bParkActive THEN
		nStep := 30;
		nCycles := 0;
	ELSIF nCycles > 10 THEN
		AssertTrue(Condition := FALSE, Message := 'the park input edge did not start the park');
		F_Note(bFailed := TRUE, sText := CONCAT(sTest, 'the park input edge did not start the park'));
		nStep := 99;
		TEST_FINISHED();
	END_IF
30:
	IF rig.fbTel.bIsParked THEN
		nStep := 40;
		nCycles := 0;
	ELSIF nCycles > 3000 THEN
		AssertTrue(Condition := FALSE, Message := 'the park did not finish');
		F_Note(bFailed := TRUE, sText := CONCAT(sTest, 'the park did not finish'));
		nStep := 99;
		TEST_FINISHED();
	END_IF
40:	// the park ended with the input still TRUE: it is not replayed and not cleared
	IF nCycles >= 30 THEN
		AssertTrue(Condition := NOT rig.fbTel.bParkActive, Message := 'the park request ended');
		F_Note(bFailed := NOT (NOT rig.fbTel.bParkActive), sText := CONCAT(sTest, 'the park request ended'));
		AssertTrue(Condition := rig.fbTel.bIsParked, Message := 'the telescope stays parked');
		F_Note(bFailed := NOT (rig.fbTel.bIsParked), sText := CONCAT(sTest, 'the telescope stays parked'));
		AssertTrue(Condition := rig.fbTel.bPark, Message := 'the block did not clear the input');
		F_Note(bFailed := NOT (rig.fbTel.bPark), sText := CONCAT(sTest, 'the block did not clear the input'));
		nStep := 99;
		TEST_FINISHED();
	END_IF
END_CASE
END_METHOD

// Stop() and a stop input edge in one scan are one command (the method sets the edge memory).
METHOD PRIVATE Stop_Method_And_Input_Edge_In_One_Scan_Count_Once
VAR_INST
	rig			: FB_IagRig;
	nStep		: INT;
	nCycles		: UINT;
	nEdges		: UINT;
	sTest		: STRING(80);
END_VAR
TEST('Stop_Method_And_Input_Edge_In_One_Scan_Count_Once');
sTest := 'Stop_Method_And_Input_Edge_In_One_Scan_Count_Once: ';
IF nStep >= 90 THEN
	RETURN;
END_IF
rig.Scan();
nCycles := nCycles + 1;
CASE nStep OF
0:	// wait for the clock, then power on
	IF rig.ClockValid THEN
		rig.fbTel.Init();
		nStep := 10;
		nCycles := 0;
	ELSIF nCycles > 2000 THEN
		AssertTrue(Condition := FALSE, Message := 'the astronomical clock never became valid');
		F_Note(bFailed := TRUE, sText := CONCAT(sTest, 'the astronomical clock never became valid'));
		nStep := 99;
		TEST_FINISHED();
	END_IF
10:	// wait until the startup has finished (READY_STATE 1.0)
	IF rig.Online THEN
		rig.fbTel.Slew(fAzimuth := 180.0, fAltitude := 45.0);
		nStep := 20;
		nCycles := 0;
	ELSIF nCycles > 1500 THEN
		AssertTrue(Condition := FALSE, Message := 'the mock telescope did not reach READY_STATE 1.0');
		F_Note(bFailed := TRUE, sText := CONCAT(sTest, 'the mock telescope did not reach READY_STATE 1.0'));
		nStep := 99;
		TEST_FINISHED();
	END_IF
20:	// an axis is moving
	IF rig.fbHa.MoveAxis OR rig.fbDec.MoveAxis THEN
		nCycles := 0;
		nStep := 30;
	ELSIF nCycles > 300 THEN
		AssertTrue(Condition := FALSE, Message := 'the slew did not start an axis move');
		F_Note(bFailed := TRUE, sText := CONCAT(sTest, 'the slew did not start an axis move'));
		nStep := 99;
		TEST_FINISHED();
	END_IF
30:	// Stop() and the input edge in the same scan
	IF nCycles >= 5 THEN
		rig.fbTel.Stop();
		rig.SetStopInput(TRUE);
		nStep := 40;
		nCycles := 0;
	END_IF
40:
	IF NOT rig.fbTel.bStopActive AND rig.fbTel.bStopped AND nCycles > 5 THEN
		AssertTrue(Condition := rig.fbFocus.nStop = 1, Message := 'one Stop(): the focus stopped once');
		F_Note(bFailed := NOT (rig.fbFocus.nStop = 1), sText := CONCAT(sTest, 'one Stop(): the focus stopped once'));
		AssertTrue(Condition := rig.fbHa.nStopEdges + rig.fbDec.nStopEdges = 1, Message := 'one stop for the moving axis');
		F_Note(bFailed := NOT (rig.fbHa.nStopEdges + rig.fbDec.nStopEdges = 1), sText := CONCAT(sTest, 'one stop for the moving axis'));
		nStep := 99;
		TEST_FINISHED();
	ELSIF nCycles > 400 THEN
		AssertTrue(Condition := FALSE, Message := 'the stop did not settle');
		F_Note(bFailed := TRUE, sText := CONCAT(sTest, 'the stop did not settle'));
		nStep := 99;
		TEST_FINISHED();
	END_IF
END_CASE
END_METHOD

// A rising power input is an Init(); the block neither clears the input nor repeats the request.
METHOD PRIVATE Power_Input_Is_Not_Written_By_The_Block
VAR_INST
	rig			: FB_IagRig;
	nStep		: INT;
	nCycles		: UINT;
	nEdges		: UINT;
	sTest		: STRING(80);
END_VAR
TEST('Power_Input_Is_Not_Written_By_The_Block');
sTest := 'Power_Input_Is_Not_Written_By_The_Block: ';
IF nStep >= 90 THEN
	RETURN;
END_IF
rig.Scan();
nCycles := nCycles + 1;
CASE nStep OF
0:	// wait for the clock, then power on
	IF rig.ClockValid THEN
		rig.SetPowerInput(TRUE);
		nStep := 10;
		nCycles := 0;
	ELSIF nCycles > 2000 THEN
		AssertTrue(Condition := FALSE, Message := 'the astronomical clock never became valid');
		F_Note(bFailed := TRUE, sText := CONCAT(sTest, 'the astronomical clock never became valid'));
		nStep := 99;
		TEST_FINISHED();
	END_IF
10:	// wait until the startup has finished (READY_STATE 1.0)
	IF rig.Online THEN
		nStep := 20;
		nCycles := 0;
	ELSIF nCycles > 1500 THEN
		AssertTrue(Condition := FALSE, Message := 'the mock telescope did not reach READY_STATE 1.0');
		F_Note(bFailed := TRUE, sText := CONCAT(sTest, 'the mock telescope did not reach READY_STATE 1.0'));
		nStep := 99;
		TEST_FINISHED();
	END_IF
20:	// the power-on ran from the input edge and finished: the latch is down, the input is what the writer left
	IF nCycles >= 30 THEN
		AssertTrue(Condition := rig.Online, Message := 'the telescope is online');
		F_Note(bFailed := NOT (rig.Online), sText := CONCAT(sTest, 'the telescope is online'));
		AssertTrue(Condition := NOT rig.fbTel.bPowerActive, Message := 'the power-on request ended');
		F_Note(bFailed := NOT (NOT rig.fbTel.bPowerActive), sText := CONCAT(sTest, 'the power-on request ended'));
		AssertTrue(Condition := rig.fbTel.bPower, Message := 'the block did not clear the input');
		F_Note(bFailed := NOT (rig.fbTel.bPower), sText := CONCAT(sTest, 'the block did not clear the input'));
		nStep := 99;
		TEST_FINISHED();
	END_IF
END_CASE
END_METHOD

// A held slew input is one slew: it runs once and is neither repeated nor cleared by the block (command model step 1b).
METHOD PRIVATE Held_Slew_Input_Starts_The_Slew_Once
VAR_INST
	rig			: FB_IagRig;
	nStep		: INT;
	nCycles		: UINT;
	nEdges		: UINT;
	sTest		: STRING(80);
END_VAR
TEST('Held_Slew_Input_Starts_The_Slew_Once');
sTest := 'Held_Slew_Input_Starts_The_Slew_Once: ';
IF nStep >= 90 THEN
	RETURN;
END_IF
rig.Scan();
nCycles := nCycles + 1;
CASE nStep OF
0:	// wait for the clock, then power on
	IF rig.ClockValid THEN
		rig.fbTel.Init();
		nStep := 10;
		nCycles := 0;
	ELSIF nCycles > 2000 THEN
		AssertTrue(Condition := FALSE, Message := 'the astronomical clock never became valid');
		F_Note(bFailed := TRUE, sText := CONCAT(sTest, 'the astronomical clock never became valid'));
		nStep := 99;
		TEST_FINISHED();
	END_IF
10:	// wait until the startup has finished (READY_STATE 1.0)
	IF rig.Online THEN
		rig.SetSlewTargetInput(180.0, 45.0);
		rig.SetSlewInput(TRUE);
		nStep := 20;
		nCycles := 0;
	ELSIF nCycles > 1500 THEN
		AssertTrue(Condition := FALSE, Message := 'the mock telescope did not reach READY_STATE 1.0');
		F_Note(bFailed := TRUE, sText := CONCAT(sTest, 'the mock telescope did not reach READY_STATE 1.0'));
		nStep := 99;
		TEST_FINISHED();
	END_IF
20:	// an axis is moving
	IF rig.fbHa.MoveAxis OR rig.fbDec.MoveAxis THEN
		nCycles := 0;
		nStep := 30;
	ELSIF nCycles > 300 THEN
		AssertTrue(Condition := FALSE, Message := 'the slew did not start an axis move');
		F_Note(bFailed := TRUE, sText := CONCAT(sTest, 'the slew did not start an axis move'));
		nStep := 99;
		TEST_FINISHED();
	END_IF
30:	// the slew from the held input runs to its end
	IF NOT rig.fbTel.bSlewActive AND rig.fbTel.bStopped AND nCycles > 5 THEN
		nStep := 40;
		nCycles := 0;
	ELSIF nCycles > 3000 THEN
		AssertTrue(Condition := FALSE, Message := 'the slew did not finish');
		F_Note(bFailed := TRUE, sText := CONCAT(sTest, 'the slew did not finish'));
		nStep := 99;
		TEST_FINISHED();
	END_IF
40:	// 60 scans with the input still TRUE: the slew is not started again, the input is not cleared
	IF nCycles >= 60 THEN
		AssertTrue(Condition := NOT rig.fbTel.bSlewActive, Message := 'the slew was not restarted');
		F_Note(bFailed := NOT (NOT rig.fbTel.bSlewActive), sText := CONCAT(sTest, 'the slew was not restarted'));
		AssertTrue(Condition := rig.fbTel.TCS_command <> E_TCSCommand.slew, Message := 'no slew command is running');
		F_Note(bFailed := NOT (rig.fbTel.TCS_command <> E_TCSCommand.slew), sText := CONCAT(sTest, 'no slew command is running'));
		AssertTrue(Condition := rig.fbTel.bSlew, Message := 'the block did not clear the input');
		F_Note(bFailed := NOT (rig.fbTel.bSlew), sText := CONCAT(sTest, 'the block did not clear the input'));
		nStep := 99;
		TEST_FINISHED();
	END_IF
END_CASE
END_METHOD

// The slew input falling does not abort the slew; it ends only by its own completion or a stop.
METHOD PRIVATE Slew_Input_Falling_Does_Not_Abort_The_Slew
VAR_INST
	rig			: FB_IagRig;
	nStep		: INT;
	nCycles		: UINT;
	nEdges		: UINT;
	sTest		: STRING(80);
END_VAR
TEST('Slew_Input_Falling_Does_Not_Abort_The_Slew');
sTest := 'Slew_Input_Falling_Does_Not_Abort_The_Slew: ';
IF nStep >= 90 THEN
	RETURN;
END_IF
rig.Scan();
nCycles := nCycles + 1;
CASE nStep OF
0:	// wait for the clock, then power on
	IF rig.ClockValid THEN
		rig.fbTel.Init();
		nStep := 10;
		nCycles := 0;
	ELSIF nCycles > 2000 THEN
		AssertTrue(Condition := FALSE, Message := 'the astronomical clock never became valid');
		F_Note(bFailed := TRUE, sText := CONCAT(sTest, 'the astronomical clock never became valid'));
		nStep := 99;
		TEST_FINISHED();
	END_IF
10:	// wait until the startup has finished (READY_STATE 1.0)
	IF rig.Online THEN
		rig.SetSlewTargetInput(180.0, 45.0);
		rig.SetSlewInput(TRUE);
		nStep := 20;
		nCycles := 0;
	ELSIF nCycles > 1500 THEN
		AssertTrue(Condition := FALSE, Message := 'the mock telescope did not reach READY_STATE 1.0');
		F_Note(bFailed := TRUE, sText := CONCAT(sTest, 'the mock telescope did not reach READY_STATE 1.0'));
		nStep := 99;
		TEST_FINISHED();
	END_IF
20:	// an axis is moving
	IF rig.fbHa.MoveAxis OR rig.fbDec.MoveAxis THEN
		nCycles := 0;
		nStep := 25;
	ELSIF nCycles > 300 THEN
		AssertTrue(Condition := FALSE, Message := 'the slew did not start an axis move');
		F_Note(bFailed := TRUE, sText := CONCAT(sTest, 'the slew did not start an axis move'));
		nStep := 99;
		TEST_FINISHED();
	END_IF
25:	// the writer drops the input while the axis moves
	IF nCycles >= 5 THEN
		rig.SetSlewInput(FALSE);
		nStep := 30;
		nCycles := 0;
	END_IF
30:
	IF nCycles >= 5 THEN
		AssertTrue(Condition := rig.fbTel.bSlewActive, Message := 'the slew goes on after the input fell');
		F_Note(bFailed := NOT (rig.fbTel.bSlewActive), sText := CONCAT(sTest, 'the slew goes on after the input fell'));
		nStep := 40;
		nCycles := 0;
	END_IF
40:
	IF NOT rig.fbTel.bSlewActive AND rig.fbTel.bStopped AND nCycles > 5 THEN
		nStep := 99;
		TEST_FINISHED();
	ELSIF nCycles > 3000 THEN
		AssertTrue(Condition := FALSE, Message := 'the slew did not finish');
		F_Note(bFailed := TRUE, sText := CONCAT(sTest, 'the slew did not finish'));
		nStep := 99;
		TEST_FINISHED();
	END_IF
END_CASE
END_METHOD

// Slew() and a slew input edge in one scan are one slew (the method sets the edge memory).
METHOD PRIVATE Slew_Method_And_Input_Edge_In_One_Scan_Count_Once
VAR_INST
	rig			: FB_IagRig;
	nStep		: INT;
	nCycles		: UINT;
	nEdges		: UINT;
	sTest		: STRING(80);
END_VAR
TEST('Slew_Method_And_Input_Edge_In_One_Scan_Count_Once');
sTest := 'Slew_Method_And_Input_Edge_In_One_Scan_Count_Once: ';
IF nStep >= 90 THEN
	RETURN;
END_IF
rig.Scan();
nCycles := nCycles + 1;
CASE nStep OF
0:	// wait for the clock, then power on
	IF rig.ClockValid THEN
		rig.fbTel.Init();
		nStep := 10;
		nCycles := 0;
	ELSIF nCycles > 2000 THEN
		AssertTrue(Condition := FALSE, Message := 'the astronomical clock never became valid');
		F_Note(bFailed := TRUE, sText := CONCAT(sTest, 'the astronomical clock never became valid'));
		nStep := 99;
		TEST_FINISHED();
	END_IF
10:	// wait until the startup has finished (READY_STATE 1.0)
	IF rig.Online THEN
		rig.fbTel.Slew(fAzimuth := 180.0, fAltitude := 45.0);
		rig.SetSlewInput(TRUE);
		nStep := 20;
		nCycles := 0;
	ELSIF nCycles > 1500 THEN
		AssertTrue(Condition := FALSE, Message := 'the mock telescope did not reach READY_STATE 1.0');
		F_Note(bFailed := TRUE, sText := CONCAT(sTest, 'the mock telescope did not reach READY_STATE 1.0'));
		nStep := 99;
		TEST_FINISHED();
	END_IF
20:	// an axis is moving
	IF rig.fbHa.MoveAxis OR rig.fbDec.MoveAxis THEN
		nCycles := 0;
		nStep := 30;
	ELSIF nCycles > 300 THEN
		AssertTrue(Condition := FALSE, Message := 'the slew did not start an axis move');
		F_Note(bFailed := TRUE, sText := CONCAT(sTest, 'the slew did not start an axis move'));
		nStep := 99;
		TEST_FINISHED();
	END_IF
30:
	IF NOT rig.fbTel.bSlewActive AND rig.fbTel.bStopped AND nCycles > 5 THEN
		nStep := 40;
		nCycles := 0;
	ELSIF nCycles > 3000 THEN
		AssertTrue(Condition := FALSE, Message := 'the slew did not finish');
		F_Note(bFailed := TRUE, sText := CONCAT(sTest, 'the slew did not finish'));
		nStep := 99;
		TEST_FINISHED();
	END_IF
40:	IF nCycles >= 60 THEN
		AssertTrue(Condition := NOT rig.fbTel.bSlewActive, Message := 'no second slew');
		F_Note(bFailed := NOT (NOT rig.fbTel.bSlewActive), sText := CONCAT(sTest, 'no second slew'));
		AssertTrue(Condition := rig.fbHa.nStopEdges + rig.fbDec.nStopEdges = 0, Message := 'no restart stop');
		F_Note(bFailed := NOT (rig.fbHa.nStopEdges + rig.fbDec.nStopEdges = 0), sText := CONCAT(sTest, 'no restart stop'));
		nStep := 99;
		TEST_FINISHED();
	END_IF
END_CASE
END_METHOD

// D1 (template body step S1.d): a slew input edge in the scan of a new axis error is rejected at arrival (the gate sees this scan's error), not accepted and dropped silently.
METHOD PRIVATE Slew_Input_In_The_Scan_Of_A_New_Error_Is_Rejected
VAR_INST
	rig			: FB_IagRig;
	nStep		: INT;
	nCycles		: UINT;
	sTest		: STRING(80);
END_VAR
TEST('Slew_Input_In_The_Scan_Of_A_New_Error_Is_Rejected');
sTest := 'Slew_Input_In_The_Scan_Of_A_New_Error_Is_Rejected: ';
IF nStep >= 90 THEN
	RETURN;
END_IF
rig.Scan();
nCycles := nCycles + 1;
CASE nStep OF
0:	// wait for the clock, then power on
	IF rig.ClockValid THEN
		rig.fbTel.Init();
		nStep := 10;
		nCycles := 0;
	ELSIF nCycles > 2000 THEN
		AssertTrue(Condition := FALSE, Message := 'the astronomical clock never became valid');
		F_Note(bFailed := TRUE, sText := CONCAT(sTest, 'the astronomical clock never became valid'));
		nStep := 99;
		TEST_FINISHED();
	END_IF
10:	// wait until the startup has finished (READY_STATE 1.0)
	IF rig.Online THEN
		rig.SetHorizon(-90.0);
		rig.SetSafeAltitude(-90.0);
		rig.SetSlewTargetInput(fAzimuth := 180.0, fAltitude := 45.0);
		rig.InjectHaError(16#4550);
		rig.SetSlewInput(TRUE);
		nStep := 20;
		nCycles := 0;
	ELSIF nCycles > 1500 THEN
		AssertTrue(Condition := FALSE, Message := 'the mock telescope did not reach READY_STATE 1.0');
		F_Note(bFailed := TRUE, sText := CONCAT(sTest, 'the mock telescope did not reach READY_STATE 1.0'));
		nStep := 99;
		TEST_FINISHED();
	END_IF
20:	// the slew edge came in the scan in which the axis error appeared: rejected at arrival, with a log, nothing latched
	IF nCycles >= 5 THEN
		AssertTrue(Condition := rig.fbTel.bError, Message := 'the error is reported');
		F_Note(bFailed := NOT (rig.fbTel.bError), sText := CONCAT(sTest, 'the error is reported'));
		AssertTrue(Condition := rig.fbTel.nCommandRejectCount >= 1, Message := 'the slew was rejected and counted');
		F_Note(bFailed := NOT (rig.fbTel.nCommandRejectCount >= 1), sText := CONCAT(sTest, 'the slew was rejected and counted'));
		AssertTrue(Condition := NOT rig.fbTel.bSlewActive, Message := 'no slew is latched');
		F_Note(bFailed := NOT (NOT rig.fbTel.bSlewActive), sText := CONCAT(sTest, 'no slew is latched'));
		nStep := 99;
		TEST_FINISHED();
	END_IF
END_CASE
END_METHOD

// D4 (template body step S1.f): Track() and a bTrack input edge in one scan are one command (Track() marks the edge memory of the track input), as in MONETcommon.
METHOD PRIVATE Track_Method_And_Track_Input_In_One_Scan_Count_Once
VAR_INST
	rig			: FB_IagRig;
	nStep		: INT;
	nCycles		: UINT;
	sTest		: STRING(80);
END_VAR
TEST('Track_Method_And_Track_Input_In_One_Scan_Count_Once');
sTest := 'Track_Method_And_Track_Input_In_One_Scan_Count_Once: ';
IF nStep >= 90 THEN
	RETURN;
END_IF
rig.Scan();
nCycles := nCycles + 1;
CASE nStep OF
0:	// wait for the clock, then power on
	IF rig.ClockValid THEN
		rig.fbTel.Init();
		nStep := 10;
		nCycles := 0;
	ELSIF nCycles > 2000 THEN
		AssertTrue(Condition := FALSE, Message := 'the astronomical clock never became valid');
		F_Note(bFailed := TRUE, sText := CONCAT(sTest, 'the astronomical clock never became valid'));
		nStep := 99;
		TEST_FINISHED();
	END_IF
10:	// wait until the startup has finished (READY_STATE 1.0)
	IF rig.Online THEN
		rig.SetHorizon(-90.0);
		rig.SetSafeAltitude(-90.0);
		rig.fbTel.Track(fRightAscension := 100.0, fDeclination := 30.0);
		rig.SetTrackInput(TRUE);
		nStep := 20;
		nCycles := 0;
	ELSIF nCycles > 1500 THEN
		AssertTrue(Condition := FALSE, Message := 'the mock telescope did not reach READY_STATE 1.0');
		F_Note(bFailed := TRUE, sText := CONCAT(sTest, 'the mock telescope did not reach READY_STATE 1.0'));
		nStep := 99;
		TEST_FINISHED();
	END_IF
20:	// one command: the goto of Track() runs, the bTrack edge of the same scan is not a second (replacing) command
	IF nCycles = 3 THEN
		AssertTrue(Condition := rig.fbTel.bGotoActive, Message := 'the goto of Track() is latched');
		F_Note(bFailed := NOT (rig.fbTel.bGotoActive), sText := CONCAT(sTest, 'the goto of Track() is latched'));
		AssertTrue(Condition := NOT rig.fbTel.bTrackActive, Message := 'the input edge did not replace it');
		F_Note(bFailed := NOT (NOT rig.fbTel.bTrackActive), sText := CONCAT(sTest, 'the input edge did not replace it'));
		AssertTrue(Condition := rig.fbTel.nCommandRejectCount = 0, Message := 'nothing was rejected');
		F_Note(bFailed := NOT (rig.fbTel.nCommandRejectCount = 0), sText := CONCAT(sTest, 'nothing was rejected'));
		AssertTrue(Condition := NOT rig.fbTel.bMoveAbortPending, Message := 'no abort stop for a replacement');
		F_Note(bFailed := NOT (NOT rig.fbTel.bMoveAbortPending), sText := CONCAT(sTest, 'no abort stop for a replacement'));
		nStep := 99;
		TEST_FINISHED();
	END_IF
END_CASE
END_METHOD

END_FUNCTION_BLOCK

// ---- POUs/IagCommandAcceptance_Tests.TcPOU
// Command acceptance at arrival (BROTLib.F_CommandAcceptance, as MONETcommon#83) in FB_TelescopeControl (IAG50cm): a move command
// that the table rejects is logged and counted and writes nothing. Plan: BROTLib specs/plans/2026-11-09-iag50cm-command-model-unification.md,
// step 2. One rig per test, one Scan() per PLC cycle.
FUNCTION_BLOCK IagCommandAcceptance_Tests EXTENDS TcUnit.FB_TestSuite
VAR
END_VAR

Slew_While_Parked_Is_Rejected();
Rejected_Slew_Writes_No_Target();
Track_During_PowerOn_Is_Rejected();
Home_While_Not_Ready_Is_Rejected();
Slew_During_Park_Is_Rejected();
Goto_During_GoHome_Is_Rejected();
Slew_During_Stop_Is_Rejected();
Rejections_Are_Counted_Each_Time();
Park_Is_Never_Rejected();

// A slew while the telescope is parked is rejected (D2), nothing is latched.
METHOD PRIVATE Slew_While_Parked_Is_Rejected
VAR_INST
	rig			: FB_IagRig;
	nStep		: INT;
	nCycles		: UINT;
	fAz			: LREAL;
	fEl			: LREAL;
	sTest		: STRING(80);
END_VAR
TEST('Slew_While_Parked_Is_Rejected');
sTest := 'Slew_While_Parked_Is_Rejected: ';
IF nStep >= 90 THEN
	RETURN;
END_IF
rig.Scan();
nCycles := nCycles + 1;
CASE nStep OF
0:	// wait for the clock, then power on
	IF rig.ClockValid THEN
		rig.fbTel.Init();
		nStep := 10;
		nCycles := 0;
	ELSIF nCycles > 2000 THEN
		AssertTrue(Condition := FALSE, Message := 'the astronomical clock never became valid');
		F_Note(bFailed := TRUE, sText := CONCAT(sTest, 'the astronomical clock never became valid'));
		nStep := 99;
		TEST_FINISHED();
	END_IF
10:	// wait until the startup has finished (READY_STATE 1.0)
	IF rig.Online THEN
		rig.fbTel.Park();
		nStep := 20;
		nCycles := 0;
	ELSIF nCycles > 1500 THEN
		AssertTrue(Condition := FALSE, Message := 'the mock telescope did not reach READY_STATE 1.0');
		F_Note(bFailed := TRUE, sText := CONCAT(sTest, 'the mock telescope did not reach READY_STATE 1.0'));
		nStep := 99;
		TEST_FINISHED();
	END_IF
20:	// wait until the park has finished
	IF rig.fbTel.bIsParked THEN
		fAz := rig.fbTel.fAzimuth;
		fEl := rig.fbTel.fElevation;
		rig.fbTel.Slew(fAzimuth := 100.0, fAltitude := 30.0);
		nStep := 30;
		nCycles := 0;
	ELSIF nCycles > 3000 THEN
		AssertTrue(Condition := FALSE, Message := 'the park did not finish');
		F_Note(bFailed := TRUE, sText := CONCAT(sTest, 'the park did not finish'));
		nStep := 99;
		TEST_FINISHED();
	END_IF
30:
		AssertTrue(Condition := rig.fbTel.nCommandRejectCount = 1, Message := 'the command was rejected and counted');
		F_Note(bFailed := NOT (rig.fbTel.nCommandRejectCount = 1), sText := CONCAT(sTest, 'the command was rejected and counted'));
		AssertTrue(Condition := rig.fbTel.eLastRejectReason = BROTLib.E_CommandRejectReason.parked, Message := 'rejected for the right reason');
		F_Note(bFailed := NOT (rig.fbTel.eLastRejectReason = BROTLib.E_CommandRejectReason.parked), sText := CONCAT(sTest, 'rejected for the right reason'));
		AssertTrue(Condition := NOT rig.fbTel.bSlewActive, Message := 'no slew was latched');
		F_Note(bFailed := NOT (NOT rig.fbTel.bSlewActive), sText := CONCAT(sTest, 'no slew was latched'));
		nStep := 99;
		TEST_FINISHED();
END_CASE
END_METHOD

// A rejected slew writes nothing, not even the target fields.
METHOD PRIVATE Rejected_Slew_Writes_No_Target
VAR_INST
	rig			: FB_IagRig;
	nStep		: INT;
	nCycles		: UINT;
	fAz			: LREAL;
	fEl			: LREAL;
	sTest		: STRING(80);
END_VAR
TEST('Rejected_Slew_Writes_No_Target');
sTest := 'Rejected_Slew_Writes_No_Target: ';
IF nStep >= 90 THEN
	RETURN;
END_IF
rig.Scan();
nCycles := nCycles + 1;
CASE nStep OF
0:	// wait for the clock, then power on
	IF rig.ClockValid THEN
		rig.fbTel.Init();
		nStep := 10;
		nCycles := 0;
	ELSIF nCycles > 2000 THEN
		AssertTrue(Condition := FALSE, Message := 'the astronomical clock never became valid');
		F_Note(bFailed := TRUE, sText := CONCAT(sTest, 'the astronomical clock never became valid'));
		nStep := 99;
		TEST_FINISHED();
	END_IF
10:	// wait until the startup has finished (READY_STATE 1.0)
	IF rig.Online THEN
		rig.fbTel.Park();
		nStep := 20;
		nCycles := 0;
	ELSIF nCycles > 1500 THEN
		AssertTrue(Condition := FALSE, Message := 'the mock telescope did not reach READY_STATE 1.0');
		F_Note(bFailed := TRUE, sText := CONCAT(sTest, 'the mock telescope did not reach READY_STATE 1.0'));
		nStep := 99;
		TEST_FINISHED();
	END_IF
20:	// wait until the park has finished
	IF rig.fbTel.bIsParked THEN
		fAz := rig.fbTel.fAzimuth;
		fEl := rig.fbTel.fElevation;
		rig.fbTel.Slew(fAzimuth := 100.0, fAltitude := 30.0);
		nStep := 30;
		nCycles := 0;
	ELSIF nCycles > 3000 THEN
		AssertTrue(Condition := FALSE, Message := 'the park did not finish');
		F_Note(bFailed := TRUE, sText := CONCAT(sTest, 'the park did not finish'));
		nStep := 99;
		TEST_FINISHED();
	END_IF
30:
		AssertTrue(Condition := rig.fbTel.nCommandRejectCount = 1, Message := 'the command was rejected and counted');
		F_Note(bFailed := NOT (rig.fbTel.nCommandRejectCount = 1), sText := CONCAT(sTest, 'the command was rejected and counted'));
		AssertTrue(Condition := rig.fbTel.eLastRejectReason = BROTLib.E_CommandRejectReason.parked, Message := 'rejected for the right reason');
		F_Note(bFailed := NOT (rig.fbTel.eLastRejectReason = BROTLib.E_CommandRejectReason.parked), sText := CONCAT(sTest, 'rejected for the right reason'));
		AssertTrue(Condition := rig.fbTel.fAzimuth = fAz AND rig.fbTel.fElevation = fEl, Message := 'the slew target is untouched');
		F_Note(bFailed := NOT (rig.fbTel.fAzimuth = fAz AND rig.fbTel.fElevation = fEl), sText := CONCAT(sTest, 'the slew target is untouched'));
		nStep := 99;
		TEST_FINISHED();
END_CASE
END_METHOD

// A track while the power-on runs is rejected (D2).
METHOD PRIVATE Track_During_PowerOn_Is_Rejected
VAR_INST
	rig			: FB_IagRig;
	nStep		: INT;
	nCycles		: UINT;
	fAz			: LREAL;
	fEl			: LREAL;
	sTest		: STRING(80);
END_VAR
TEST('Track_During_PowerOn_Is_Rejected');
sTest := 'Track_During_PowerOn_Is_Rejected: ';
IF nStep >= 90 THEN
	RETURN;
END_IF
rig.Scan();
nCycles := nCycles + 1;
CASE nStep OF
0:	// wait for the clock
	IF rig.ClockValid THEN
		rig.fbTel.Init();
		nStep := 10;
		nCycles := 0;
	ELSIF nCycles > 2000 THEN
		AssertTrue(Condition := FALSE, Message := 'the astronomical clock never became valid');
		F_Note(bFailed := TRUE, sText := CONCAT(sTest, 'the astronomical clock never became valid'));
		nStep := 99;
		TEST_FINISHED();
	END_IF
10:	// the power-on is running
	rig.fbTel.Track(fRightAscension := 100.0, fDeclination := 30.0);
	nStep := 20;
20:
		AssertTrue(Condition := rig.fbTel.nCommandRejectCount = 1, Message := 'the command was rejected and counted');
		F_Note(bFailed := NOT (rig.fbTel.nCommandRejectCount = 1), sText := CONCAT(sTest, 'the command was rejected and counted'));
		AssertTrue(Condition := rig.fbTel.eLastRejectReason = BROTLib.E_CommandRejectReason.powering_on, Message := 'rejected for the right reason');
		F_Note(bFailed := NOT (rig.fbTel.eLastRejectReason = BROTLib.E_CommandRejectReason.powering_on), sText := CONCAT(sTest, 'rejected for the right reason'));
		AssertTrue(Condition := NOT rig.fbTel.bGotoActive, Message := 'no goto was latched');
		F_Note(bFailed := NOT (NOT rig.fbTel.bGotoActive), sText := CONCAT(sTest, 'no goto was latched'));
		nStep := 99;
		TEST_FINISHED();
END_CASE
END_METHOD

// A home while the telescope is not ready is rejected, not left pending for 2 minutes (D4).
METHOD PRIVATE Home_While_Not_Ready_Is_Rejected
VAR_INST
	rig			: FB_IagRig;
	nStep		: INT;
	nCycles		: UINT;
	fAz			: LREAL;
	fEl			: LREAL;
	sTest		: STRING(80);
END_VAR
TEST('Home_While_Not_Ready_Is_Rejected');
sTest := 'Home_While_Not_Ready_Is_Rejected: ';
IF nStep >= 90 THEN
	RETURN;
END_IF
rig.Scan();
nCycles := nCycles + 1;
CASE nStep OF
0:	// wait for the clock
	IF rig.ClockValid THEN
		rig.fbTel.Home();
		nStep := 10;
		nCycles := 0;
	ELSIF nCycles > 2000 THEN
		AssertTrue(Condition := FALSE, Message := 'the astronomical clock never became valid');
		F_Note(bFailed := TRUE, sText := CONCAT(sTest, 'the astronomical clock never became valid'));
		nStep := 99;
		TEST_FINISHED();
	END_IF
10:
		AssertTrue(Condition := rig.fbTel.nCommandRejectCount = 1, Message := 'the home was rejected and counted');
		F_Note(bFailed := NOT (rig.fbTel.nCommandRejectCount = 1), sText := CONCAT(sTest, 'the home was rejected and counted'));
		AssertTrue(Condition := rig.fbTel.eLastRejectReason <> BROTLib.E_CommandRejectReason.none, Message := 'with a reason');
		F_Note(bFailed := NOT (rig.fbTel.eLastRejectReason <> BROTLib.E_CommandRejectReason.none), sText := CONCAT(sTest, 'with a reason'));
		AssertTrue(Condition := NOT rig.fbTel.bGoHomeActive, Message := 'no home was latched (it used to wait 2 min)');
		F_Note(bFailed := NOT (NOT rig.fbTel.bGoHomeActive), sText := CONCAT(sTest, 'no home was latched (it used to wait 2 min)'));
		nStep := 99;
		TEST_FINISHED();
END_CASE
END_METHOD

// A slew while a park is pending or running is rejected (D2).
METHOD PRIVATE Slew_During_Park_Is_Rejected
VAR_INST
	rig			: FB_IagRig;
	nStep		: INT;
	nCycles		: UINT;
	fAz			: LREAL;
	fEl			: LREAL;
	sTest		: STRING(80);
END_VAR
TEST('Slew_During_Park_Is_Rejected');
sTest := 'Slew_During_Park_Is_Rejected: ';
IF nStep >= 90 THEN
	RETURN;
END_IF
rig.Scan();
nCycles := nCycles + 1;
CASE nStep OF
0:	// wait for the clock, then power on
	IF rig.ClockValid THEN
		rig.fbTel.Init();
		nStep := 10;
		nCycles := 0;
	ELSIF nCycles > 2000 THEN
		AssertTrue(Condition := FALSE, Message := 'the astronomical clock never became valid');
		F_Note(bFailed := TRUE, sText := CONCAT(sTest, 'the astronomical clock never became valid'));
		nStep := 99;
		TEST_FINISHED();
	END_IF
10:	// wait until the startup has finished (READY_STATE 1.0)
	IF rig.Online THEN
		rig.fbTel.Park();
		nStep := 20;
		nCycles := 0;
	ELSIF nCycles > 1500 THEN
		AssertTrue(Condition := FALSE, Message := 'the mock telescope did not reach READY_STATE 1.0');
		F_Note(bFailed := TRUE, sText := CONCAT(sTest, 'the mock telescope did not reach READY_STATE 1.0'));
		nStep := 99;
		TEST_FINISHED();
	END_IF
20:	// the park is running
	IF rig.fbTel.bParkActive THEN
		rig.fbTel.Slew(fAzimuth := 100.0, fAltitude := 30.0);
		nStep := 30;
		nCycles := 0;
	ELSIF nCycles > 10 THEN
		AssertTrue(Condition := FALSE, Message := 'the park did not start');
		F_Note(bFailed := TRUE, sText := CONCAT(sTest, 'the park did not start'));
		nStep := 99;
		TEST_FINISHED();
	END_IF
30:
		AssertTrue(Condition := rig.fbTel.nCommandRejectCount = 1, Message := 'the command was rejected and counted');
		F_Note(bFailed := NOT (rig.fbTel.nCommandRejectCount = 1), sText := CONCAT(sTest, 'the command was rejected and counted'));
		AssertTrue(Condition := rig.fbTel.eLastRejectReason = BROTLib.E_CommandRejectReason.parking, Message := 'rejected for the right reason');
		F_Note(bFailed := NOT (rig.fbTel.eLastRejectReason = BROTLib.E_CommandRejectReason.parking), sText := CONCAT(sTest, 'rejected for the right reason'));
		nStep := 99;
		TEST_FINISHED();
END_CASE
END_METHOD

// A goto/track while the home runs is rejected (D2).
METHOD PRIVATE Goto_During_GoHome_Is_Rejected
VAR_INST
	rig			: FB_IagRig;
	nStep		: INT;
	nCycles		: UINT;
	fAz			: LREAL;
	fEl			: LREAL;
	sTest		: STRING(80);
END_VAR
TEST('Goto_During_GoHome_Is_Rejected');
sTest := 'Goto_During_GoHome_Is_Rejected: ';
IF nStep >= 90 THEN
	RETURN;
END_IF
rig.Scan();
nCycles := nCycles + 1;
CASE nStep OF
0:	// wait for the clock, then power on
	IF rig.ClockValid THEN
		rig.fbTel.Init();
		nStep := 10;
		nCycles := 0;
	ELSIF nCycles > 2000 THEN
		AssertTrue(Condition := FALSE, Message := 'the astronomical clock never became valid');
		F_Note(bFailed := TRUE, sText := CONCAT(sTest, 'the astronomical clock never became valid'));
		nStep := 99;
		TEST_FINISHED();
	END_IF
10:	// wait until the startup has finished (READY_STATE 1.0)
	IF rig.Online THEN
		rig.fbTel.Home();
		nStep := 20;
		nCycles := 0;
	ELSIF nCycles > 1500 THEN
		AssertTrue(Condition := FALSE, Message := 'the mock telescope did not reach READY_STATE 1.0');
		F_Note(bFailed := TRUE, sText := CONCAT(sTest, 'the mock telescope did not reach READY_STATE 1.0'));
		nStep := 99;
		TEST_FINISHED();
	END_IF
20:	// the home is accepted and running
	IF rig.fbTel.bGoHomeActive THEN
		AssertTrue(Condition := rig.fbTel.nCommandRejectCount = 0, Message := 'the home from the ready telescope was accepted');
		F_Note(bFailed := NOT (rig.fbTel.nCommandRejectCount = 0), sText := CONCAT(sTest, 'the home from the ready telescope was accepted'));
		rig.fbTel.Track(fRightAscension := 100.0, fDeclination := 30.0);
		nStep := 30;
		nCycles := 0;
	ELSIF nCycles > 10 THEN
		AssertTrue(Condition := FALSE, Message := 'the home did not start');
		F_Note(bFailed := TRUE, sText := CONCAT(sTest, 'the home did not start'));
		nStep := 99;
		TEST_FINISHED();
	END_IF
30:
		AssertTrue(Condition := rig.fbTel.nCommandRejectCount = 1, Message := 'the command was rejected and counted');
		F_Note(bFailed := NOT (rig.fbTel.nCommandRejectCount = 1), sText := CONCAT(sTest, 'the command was rejected and counted'));
		AssertTrue(Condition := rig.fbTel.eLastRejectReason = BROTLib.E_CommandRejectReason.gohome_active, Message := 'rejected for the right reason');
		F_Note(bFailed := NOT (rig.fbTel.eLastRejectReason = BROTLib.E_CommandRejectReason.gohome_active), sText := CONCAT(sTest, 'rejected for the right reason'));
		nStep := 99;
		TEST_FINISHED();
END_CASE
END_METHOD

// A slew while a stop is running is rejected (D5).
METHOD PRIVATE Slew_During_Stop_Is_Rejected
VAR_INST
	rig			: FB_IagRig;
	nStep		: INT;
	nCycles		: UINT;
	fAz			: LREAL;
	fEl			: LREAL;
	sTest		: STRING(80);
END_VAR
TEST('Slew_During_Stop_Is_Rejected');
sTest := 'Slew_During_Stop_Is_Rejected: ';
IF nStep >= 90 THEN
	RETURN;
END_IF
rig.Scan();
nCycles := nCycles + 1;
CASE nStep OF
0:	// wait for the clock, then power on
	IF rig.ClockValid THEN
		rig.fbTel.Init();
		nStep := 10;
		nCycles := 0;
	ELSIF nCycles > 2000 THEN
		AssertTrue(Condition := FALSE, Message := 'the astronomical clock never became valid');
		F_Note(bFailed := TRUE, sText := CONCAT(sTest, 'the astronomical clock never became valid'));
		nStep := 99;
		TEST_FINISHED();
	END_IF
10:	// wait until the startup has finished (READY_STATE 1.0)
	IF rig.Online THEN
		rig.fbTel.Slew(fAzimuth := 180.0, fAltitude := 45.0);
		nStep := 20;
		nCycles := 0;
	ELSIF nCycles > 1500 THEN
		AssertTrue(Condition := FALSE, Message := 'the mock telescope did not reach READY_STATE 1.0');
		F_Note(bFailed := TRUE, sText := CONCAT(sTest, 'the mock telescope did not reach READY_STATE 1.0'));
		nStep := 99;
		TEST_FINISHED();
	END_IF
20:	// an axis is moving: stop
	IF rig.fbHa.MoveAxis OR rig.fbDec.MoveAxis THEN
		rig.fbTel.Stop();
		nStep := 30;
		nCycles := 0;
	ELSIF nCycles > 300 THEN
		AssertTrue(Condition := FALSE, Message := 'the slew did not start an axis move');
		F_Note(bFailed := TRUE, sText := CONCAT(sTest, 'the slew did not start an axis move'));
		nStep := 99;
		TEST_FINISHED();
	END_IF
30:	// the stop is running
	IF rig.fbTel.bStopActive THEN
		rig.fbTel.Slew(fAzimuth := 100.0, fAltitude := 30.0);
		nStep := 40;
		nCycles := 0;
	ELSIF nCycles > 10 THEN
		AssertTrue(Condition := FALSE, Message := 'the stop did not start');
		F_Note(bFailed := TRUE, sText := CONCAT(sTest, 'the stop did not start'));
		nStep := 99;
		TEST_FINISHED();
	END_IF
40:
		AssertTrue(Condition := rig.fbTel.nCommandRejectCount = 1, Message := 'the command was rejected and counted');
		F_Note(bFailed := NOT (rig.fbTel.nCommandRejectCount = 1), sText := CONCAT(sTest, 'the command was rejected and counted'));
		AssertTrue(Condition := rig.fbTel.eLastRejectReason = BROTLib.E_CommandRejectReason.stopping, Message := 'rejected for the right reason');
		F_Note(bFailed := NOT (rig.fbTel.eLastRejectReason = BROTLib.E_CommandRejectReason.stopping), sText := CONCAT(sTest, 'rejected for the right reason'));
		nStep := 99;
		TEST_FINISHED();
END_CASE
END_METHOD

// Every rejection is counted, also an identical one in consecutive scans (the log shows an identical one within 2 s once).
METHOD PRIVATE Rejections_Are_Counted_Each_Time
VAR_INST
	rig			: FB_IagRig;
	nStep		: INT;
	nCycles		: UINT;
	fAz			: LREAL;
	fEl			: LREAL;
	sTest		: STRING(80);
END_VAR
TEST('Rejections_Are_Counted_Each_Time');
sTest := 'Rejections_Are_Counted_Each_Time: ';
IF nStep >= 90 THEN
	RETURN;
END_IF
rig.Scan();
nCycles := nCycles + 1;
CASE nStep OF
0:	// wait for the clock, then power on
	IF rig.ClockValid THEN
		rig.fbTel.Init();
		nStep := 10;
		nCycles := 0;
	ELSIF nCycles > 2000 THEN
		AssertTrue(Condition := FALSE, Message := 'the astronomical clock never became valid');
		F_Note(bFailed := TRUE, sText := CONCAT(sTest, 'the astronomical clock never became valid'));
		nStep := 99;
		TEST_FINISHED();
	END_IF
10:	// wait until the startup has finished (READY_STATE 1.0)
	IF rig.Online THEN
		rig.fbTel.Park();
		nStep := 20;
		nCycles := 0;
	ELSIF nCycles > 1500 THEN
		AssertTrue(Condition := FALSE, Message := 'the mock telescope did not reach READY_STATE 1.0');
		F_Note(bFailed := TRUE, sText := CONCAT(sTest, 'the mock telescope did not reach READY_STATE 1.0'));
		nStep := 99;
		TEST_FINISHED();
	END_IF
20:
	IF rig.fbTel.bIsParked THEN
		rig.fbTel.Slew(fAzimuth := 100.0, fAltitude := 30.0);
		nStep := 30;
		nCycles := 0;
	ELSIF nCycles > 3000 THEN
		AssertTrue(Condition := FALSE, Message := 'the park did not finish');
		F_Note(bFailed := TRUE, sText := CONCAT(sTest, 'the park did not finish'));
		nStep := 99;
		TEST_FINISHED();
	END_IF
30:	// a second rejection in the next scan
	rig.fbTel.Slew(fAzimuth := 100.0, fAltitude := 30.0);
	nStep := 40;
40:
		AssertTrue(Condition := rig.fbTel.nCommandRejectCount = 2, Message := 'both rejections are counted');
		F_Note(bFailed := NOT (rig.fbTel.nCommandRejectCount = 2), sText := CONCAT(sTest, 'both rejections are counted'));
		nStep := 99;
		TEST_FINISHED();
END_CASE
END_METHOD

// A park is never rejected by the acceptance table.
METHOD PRIVATE Park_Is_Never_Rejected
VAR_INST
	rig			: FB_IagRig;
	nStep		: INT;
	nCycles		: UINT;
	fAz			: LREAL;
	fEl			: LREAL;
	sTest		: STRING(80);
END_VAR
TEST('Park_Is_Never_Rejected');
sTest := 'Park_Is_Never_Rejected: ';
IF nStep >= 90 THEN
	RETURN;
END_IF
rig.Scan();
nCycles := nCycles + 1;
CASE nStep OF
0:	// wait for the clock
	IF rig.ClockValid THEN
		rig.fbTel.Init();
		nStep := 10;
		nCycles := 0;
	ELSIF nCycles > 2000 THEN
		AssertTrue(Condition := FALSE, Message := 'the astronomical clock never became valid');
		F_Note(bFailed := TRUE, sText := CONCAT(sTest, 'the astronomical clock never became valid'));
		nStep := 99;
		TEST_FINISHED();
	END_IF
10:	// the power-on is running: a park is not rejected, it wins over the power-on
	rig.fbTel.Park();
	nStep := 20;
	nCycles := 0;
20:
	IF nCycles >= 5 THEN
		AssertTrue(Condition := rig.fbTel.nCommandRejectCount = 0, Message := 'a park is never rejected');
		F_Note(bFailed := NOT (rig.fbTel.nCommandRejectCount = 0), sText := CONCAT(sTest, 'a park is never rejected'));
		AssertTrue(Condition := rig.fbTel.bParkActive OR rig.fbTel.bIsParked, Message := 'the park runs');
		F_Note(bFailed := NOT (rig.fbTel.bParkActive OR rig.fbTel.bIsParked), sText := CONCAT(sTest, 'the park runs'));
		nStep := 99;
		TEST_FINISHED();
	END_IF
END_CASE
END_METHOD

END_FUNCTION_BLOCK

// ---- POUs/IagAbortStop_Tests.TcPOU
// Abort stop and stop semantics of FB_TelescopeControl (IAG50cm), command model step 3A (BROTLib
// specs/plans/2026-11-09-iag50cm-command-model-unification.md). One rig per test, one Scan() per PLC cycle.
FUNCTION_BLOCK IagAbortStop_Tests EXTENDS TcUnit.FB_TestSuite
VAR
END_VAR

Error_During_Abort_Stop_Clears_It();
Stop_Is_Held_Until_The_Transaction_Settles();
Stop_Clears_Every_Pending_Move();
Repeated_Stop_Restarts_Only_Moving_Axes();
Park_Over_A_Waiting_Goto_Runs_A_Short_Abort_Stop();

// An error clears the abort stop: the drives are disabled, there is nothing to wait for (3A.1).
METHOD PRIVATE Error_During_Abort_Stop_Clears_It
VAR_INST
	rig			: FB_IagRig;
	nStep		: INT;
	nCycles		: UINT;
	nEdges		: UINT;
	bSeen		: BOOL;
	sTest		: STRING(80);
END_VAR
TEST('Error_During_Abort_Stop_Clears_It');
sTest := 'Error_During_Abort_Stop_Clears_It: ';
IF nStep >= 90 THEN
	RETURN;
END_IF
rig.Scan();
nCycles := nCycles + 1;
CASE nStep OF
0:	// wait for the clock, then power on
	IF rig.ClockValid THEN
		rig.fbTel.Init();
		nStep := 10;
		nCycles := 0;
	ELSIF nCycles > 2000 THEN
		AssertTrue(Condition := FALSE, Message := 'the astronomical clock never became valid');
		F_Note(bFailed := TRUE, sText := CONCAT(sTest, 'the astronomical clock never became valid'));
		nStep := 99;
		TEST_FINISHED();
	END_IF
10:	// wait until the startup has finished (READY_STATE 1.0)
	IF rig.Online THEN
		// the target is not checked against the sky of the day this runs on: no horizon, no safe altitude
		rig.SetHorizon(-90.0);
		rig.SetSafeAltitude(-90.0);
		rig.fbTel.Track(fRightAscension := 100.0, fDeclination := 30.0);
		nStep := 20;
		nCycles := 0;
	ELSIF nCycles > 1500 THEN
		AssertTrue(Condition := FALSE, Message := 'the mock telescope did not reach READY_STATE 1.0');
		F_Note(bFailed := TRUE, sText := CONCAT(sTest, 'the mock telescope did not reach READY_STATE 1.0'));
		nStep := 99;
		TEST_FINISHED();
	END_IF
20:	// the goto runs: a second track replaces it through the abort stop
	IF rig.fbHa.MoveAxis OR rig.fbDec.MoveAxis THEN
		rig.fbTel.Track(fRightAscension := 110.0, fDeclination := 31.0);
		nStep := 25;
		nCycles := 0;
	ELSIF nCycles > 300 THEN
		AssertTrue(Condition := FALSE, Message := 'the goto did not start an axis move');
		F_Note(bFailed := TRUE, sText := CONCAT(sTest, 'the goto did not start an axis move'));
		nStep := 99;
		TEST_FINISHED();
	END_IF
25:
	IF rig.fbTel.bMoveAbortPending THEN
		rig.InjectHaError(16#4550);
		nStep := 30;
		nCycles := 0;
	ELSIF nCycles > 10 THEN
		AssertTrue(Condition := FALSE, Message := 'the replaced goto did not run an abort stop');
		F_Note(bFailed := TRUE, sText := CONCAT(sTest, 'the replaced goto did not run an abort stop'));
		nStep := 99;
		TEST_FINISHED();
	END_IF
30:
	IF nCycles >= 5 THEN
		AssertTrue(Condition := rig.fbTel.bError, Message := 'the axis error is seen');
		F_Note(bFailed := NOT (rig.fbTel.bError), sText := CONCAT(sTest, 'the axis error is seen'));
		AssertTrue(Condition := NOT rig.fbTel.bMoveAbortPending, Message := 'the error cleared the abort stop');
		F_Note(bFailed := NOT (NOT rig.fbTel.bMoveAbortPending), sText := CONCAT(sTest, 'the error cleared the abort stop'));
		nStep := 99;
		TEST_FINISHED();
	END_IF
END_CASE
END_METHOD

